Universal Robots PolyScope program: AdientTorsF_Eol20.urp

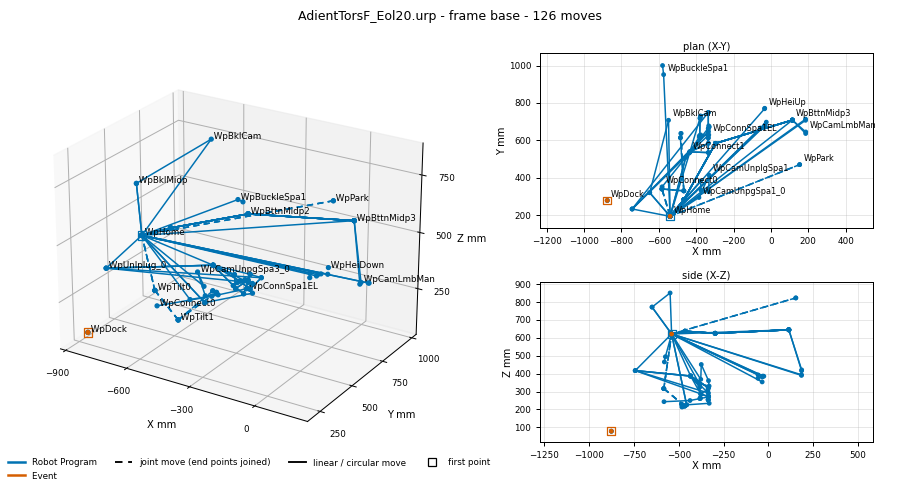
[picture p0: tool path of AdientTorsF_Eol20.urp in frame base, 126 of 179 moves have a stored position in this frame; points joined in program order, loops and branches not executed]
Program AdientTorsF_Eol20 (installation=EOL_20 directory=/programs createdIn=3.5.1 lastSavedIn=5.26.0 robotSerialNumber=20265101888)
Calibrated DH parameters: a=[0.000055, -0.599562, -0.553909, 0.000045, 0.000002, 0]; d=[0.180957, -130.68916, 109.469633, 21.394116, 0.119819, 0.115629]; alpha=[1.570664, -0.000951, 0.006615, 1.571213, -1.569974, 0]; deltaTheta=[0, 0.204436, 5.830565, 0.248193, -0.000001, 0]
InitVariablesNode variables(variable(name=Abort, expression=False), variable(name=AdapterReady, expression=False), variable(name=CMD_Heartbt_i1, expression=0), variable(name=CMD_Program_i1, expression=0), variable(name=CMD_Reserve_i1, expression=0), variable(name=CMD_Timeout_i1, expression=0), variable(name=CamCorrectnOK, expression=0), variable(name=DEBUG, expression=False), variable(name=D_rel, expression=p[0,0,0,0,0,0]), variable(name=EvtBeep, expression=False), variable(name=EvtDock, expression=0), variable(name=Mute, expression=False), variable(name=P_ini, expression=get_actual_tcp_pose()), variable(name=Parking, expression=0), variable(name=ProgExe, expression=0), variable(name=PusherPosFt, expression=0), variable(name=PusherReturn, expression=True), variable(name=STS_Heartbeat, expression=False), variable(name=STS_Progress, expression=0), variable(name=STS_Reservation, expression=0), variable(name=SetCameraProg, expression=0), variable(name=T_KeepReservtn, expression=0), variable(name=Tilt_PV, expression=0))
BeforeStart
  SuppressedNode
    DEBUG := True
  'SW version, to be used to track changes and keep sync of all stations'
  SW_Ver := 1.0
  Folder Scripts [hidden by the author, left out]
  Folder Avoid guidance screen
    Wp := get_actual_tcp_pose()
    MoveJ speed 120 deg/s, acceleration 500 deg/s^2 (useActiveTCP=true optimoveEnabled=false optiMoveSpeed=0.3 optiMoveAcceleration=0.09) feature=Base
      Waypoint Variable (Variable): variable=Wp
  Call GripperOpen
  GoToHome := True
  Script: socket_open("127.0.0.1",30001)
Robot Program (runOnlyOnce=false)
  Folder Execute Program
    Folder Init
      Wait Condition expression=EvtDock≤0
      Folder Verify Adapter ready
        If digital_in[0] or analog_in[3]<(ivGripSensOpen+0.3)
          AdapterReady := False
      Folder Go to home pos automatically
        If GoToHome and  not AdapterReady
          Wait Sleep waitTime=1
          If InRange(P_Flange[0],-1,-0.2) and InRange(P_Flange[1],-0.5,0.5) and InRange(P_Flange[2],0.3,1)
            If AdapterDocked or DEBUG or (analog_in[3]<(ivGripSensOpen+0.3))
              MoveJ speed 120 deg/s, acceleration 500 deg/s^2 (useActiveTCP=false positionType=JointAngles optimoveEnabled=false optiMoveSpeed=0.3 optiMoveAcceleration=0.09) tcp=t0_Flange; feature=Base
                Waypoint WpHome: TCP in base x=-539.74 y=192.879 z=621.496 mm, rx=3.1416 ry=0 rz=0 rad; joints [177.915, -76.399, -107.627, -86.021, 90.391, 88.106] deg
            Else 
              Popup Error (haltProgram=false message=Adapter must be docked inputType=Text)
              Halt
          ElseIf AtParkPos
            MoveJ speed 120 deg/s, acceleration 500 deg/s^2 (useActiveTCP=false positionType=JointAngles optimoveEnabled=false optiMoveSpeed=0.3 optiMoveAcceleration=0.09) tcp=t0_Flange; feature=Base
              Waypoint WpPark: TCP in base x=153.666 y=469.873 z=822.74 mm, rx=-0.0357 ry=3.1413 rz=-0.0002 rad; joints [92.418, -70.926, -90.975, -108.153, 90.407, 181.161] deg
          Else 
            Popup Error (haltProgram=false message=Illegal position. Adjust arm to open space in front of the backrest, or [Move]->[Home] inputType=Text)
            Halt
        GoToHome := False
      If DEBUG
        'Popup window with program selection'
        ProgExe :=  (valueSource=Operator message=Program number? valueType=Integer)
      If ProgExe>0
        Folder Init
          Mute := False
          Wait Condition expression=not GoToHome
          If not In(ProgExe,[11,12,13,14])
            AdapterReady := False
    Folder Programs
      If InRange(ProgExe,1,99)
        Folder Undock
          If In(ProgExe,[11])
            Script: Report(1)
            If not AdapterReady
              Folder AtHome? [hidden by the author, left out]
              If Progress_run() and  not AdapterDocked
                Script: Report(94)
              If Progress_run()
                Folder Undock
                  MoveL speed 1000 mm/s, acceleration 3000 mm/s^2 (useActiveTCP=false optimoveEnabled=false optiMoveSpeed=0.3 optiMoveAcceleration=0.09) tcp=t2_Gripper; feature=Base
                    Call GripperOpenQuick
                    Wp := pose_trans(WpDock, p[0,0.175,-0.1,0,0,0])
                    Waypoint Variable (Variable): motionParameters(blendRadius=0.05); variable=Wp
                    Call GripperOpen
                    Wp := pose_trans(WpDock, p[0,0.075,0.01,0,0,0])
                    Waypoint Variable (Variable): motionParameters(blendRadius=0.01); variable=Wp
                    Wp := pose_trans(WpDock, p[0,0.055,0,0,0,0])
                    Waypoint Variable (Variable): motionParameters(blendRadius=0.01); variable=Wp
                    Waypoint WpDock: TCP in base x=-876.296 y=277.871 z=78.699 mm, rx=1.8725 ry=1.8725 rz=0.5904 rad; joints [172.393, -110.839, -101.123, -92.857, 86.047, -6.096] deg
                    Call GripperClose
                    Wp := pose_trans(WpDock, p[0,0.25,0,0,0,0])
                    Waypoint Variable (Variable): variable=Wp
                  AdapterReady := True
                  Script: Report(50)
            Else 
              Script: Report(50)
        Folder Connect
          If In(ProgExe,[12,13,14])
            Script: Report(1)
            PusherPosDev := 0
            MeasHeight := 0
            If not AdapterReady
              Folder AtHome? [hidden by the author, left out]
              If Progress_run() and  not AdapterDocked
                Script: Report(94)
            If Progress_run()
              Folder Length measure with pusher (mechanical seat)
                If In(ProgExe,[13])
                  Set DigitalOutput pin=Do_PusherReturn; digitalValue=0
                  Set DigitalOutput pin=Do_PusherWork; digitalValue=1
                Else 
                  PusherReturn := True
              Folder Undock
                If not AdapterReady
                  MoveL speed 1000 mm/s, acceleration 3000 mm/s^2 (useActiveTCP=false optimoveEnabled=false optiMoveSpeed=0.3 optiMoveAcceleration=0.09) tcp=t2_Gripper; feature=Base
                    Call GripperOpenQuick
                    Wp := pose_trans(WpDock, p[0,0.175,-0.1,0,0,0])
                    Waypoint Variable (Variable): motionParameters(blendRadius=0.05); variable=Wp
                    Call GripperOpen
                    Wp := pose_trans(WpDock, p[0,0.075,0.01,0,0,0])
                    Waypoint Variable (Variable): motionParameters(blendRadius=0.01); variable=Wp
                    Wp := pose_trans(WpDock, p[0,0.055,0,0,0,0])
                    Waypoint Variable (Variable): motionParameters(blendRadius=0.01); variable=Wp
                    Waypoint WpDock: TCP in base x=-876.296 y=277.871 z=78.699 mm, rx=1.8725 ry=1.8725 rz=0.5904 rad; joints [172.393, -110.839, -101.123, -92.857, 86.047, -6.096] deg
                    Call GripperClose
                    Wp := pose_trans(WpDock, p[0,0.25,0,0,0,0])
                    Waypoint Variable (Variable): variable=Wp
                AdapterReady := False
                Script: Report(2)
              CamCorrection := p[0,0,0,0,0,0]
              SuppressedNode
                Folder Camera
                  MoveL speed 1000 mm/s, acceleration 3000 mm/s^2 (useActiveTCP=false optimoveEnabled=false optiMoveSpeed=0.3 optiMoveAcceleration=0.09) tcp=t0_Flange; feature=Base
                    If In(ProgExe,[12,13])
                      SetCameraProg := 12
                      Waypoint WpCamCon0: motionParameters(blendRadius=0.05); TCP in base x=-326.648 y=291.698 z=338.41 mm, rx=2.1948 ry=2.1949 rz=-0.0575 rad; joints [160.702, -71.24, -141.099, -58.684, 93.132, -18.987] deg
                      Waypoint WpCamConSpa1: TCP in base x=-326.648 y=416.698 z=338.41 mm, rx=2.1948 ry=2.1949 rz=-0.0575 rad; joints [146.583, -82.407, -133.037, -56.241, 92.784, -33.102] deg
                    If In(ProgExe,[14])
                      SetCameraProg := ProgExe
                      Waypoint WpCamCon0: motionParameters(blendRadius=0.05); TCP in base x=-326.648 y=291.698 z=338.41 mm, rx=2.1948 ry=2.1949 rz=-0.0575 rad; joints [160.702, -71.24, -141.099, -58.684, 93.132, -18.987] deg
                      Waypoint WpCamConSpa3: TCP in base x=-370.516 y=382.662 z=354.732 mm, rx=-2.2214 ry=-2.2215 rz=0 rad; joints [153.025, -81.286, -132.366, -56.394, 90.281, -26.621] deg
                  Call CamAcquire
                  CamCorrection := p[CamData[0],CamData[1]*-0.5,CamData[1],0,0,0]
            CamCorrectnOK := ProgExe
            If In(ProgExe,[13])
              Timer (action=Reset) variable=T_Timeout
              Timer (action=Start) variable=T_Timeout
              Wait Condition expression=(PusherPosStable and InRange(PusherPos-ivPusherSeatRef,-15,15)) or T_Timeout>10
              PusherPosDev := PusherPos-ivPusherSeatRef
              If PusherPosStable and InRange(PusherPosDev,-15,15)
                'continue'
              Else 
                CamCorrectnOK := 0
                'CamCorrectionOK is also used as pusher measurement result'
            If Progress_run() and CamCorrectnOK≠ProgExe
              EvtDock := 1
              Wait Condition expression=EvtDock≤0
              Script: Report(91)
            If Progress_run() and ProgExe≟13
              'Wait handle catch done'
              Script: Report(3)
              Timer (action=Reset) variable=T_Timeout
              Timer (action=Start) variable=T_Timeout
              Wait Condition expression=Flags[12] or T_Timeout>10 or DEBUG
              If Flags[12] or DEBUG
                'ok'
              Else 
                Script: Report(98)
            If Progress_run() and  not Di_LiftDown
              EvtDock := 1
              Wait Condition expression=EvtDock≤0
              AdapterReady := False
              Script: Report(92)
            Folder Connect
              If Progress_run()
                Script: Report(4)
                Set NoAction tcp=t2_Gripper
                MoveL speed 1000 mm/s, acceleration 3000 mm/s^2 (useActiveTCP=false optimoveEnabled=false optiMoveSpeed=0.3 optiMoveAcceleration=0.09) tcp=t2_Gripper; feature=Base
                  Waypoint WpConnect0: motionParameters(blendRadius=0.01); TCP in base x=-582.317 y=351.257 z=243.437 mm, rx=-2.2214 ry=-2.2215 rz=0 rad; joints [153.816, -77.664, -139.707, -52.675, 90.266, -25.814] deg; TCP offset x=0 y=-260 z=74 mm, rx=0 ry=0 rz=0 rad
                  Waypoint WpConnect1: TCP in base x=-437.091 y=531.932 z=249.935 mm, rx=3.1416 ry=0 rz=0 rad; joints [167.745, -81.605, -135.899, -52.542, 90.261, 78.118] deg
                  If False
                    Waypoint WpConnSpa1EL: TCP in base x=-332.78 y=629.084 z=270.528 mm, rx=3.1251 ry=-0.0345 rz=0.0169 rad; joints [152.504, -78.36, -135.112, -57.546, 90.839, 64.112] deg
                    Waypoint WpConnSpa1MecTh: TCP in base x=-333.346 y=677.301 z=275.481 mm, rx=3.0512 ry=-0.0001 rz=0 rad; joints [145.822, -81.498, -129.414, -62.023, 94.591, 56.042] deg
                    Waypoint WpConnSpa1Mec: TCP in base x=-335.918 y=624.072 z=312.701 mm, rx=3.0512 ry=-0.0001 rz=0 rad; joints [151.192, -74.921, -130.239, -67.362, 94.873, 61.392] deg
                    Waypoint WpConnSpa3: TCP in base x=-375.972 y=628.734 z=287.575 mm, rx=2.9708 ry=0 rz=0.0001 rad; joints [151.145, -79.992, -126.667, -68.106, 98.894, 61.08] deg
                  If In(ProgExe,[12])
                    Wp := WpConnSpa1EL
                  If In(ProgExe,[13])
                    'adjust angle mechanical'
                    Wp0 := pose_add(WpConnSpa1MecTh,p[0,PusherPosDev/1000,-0.025,0,0,0])
                    Waypoint Variable (Variable): variable=Wp0
                    Force Frame feature=Joint_6_name; selection=[0, 0, 1, 0, 0, 0]; wrench=[0, 0, -30, -0.5, 0, 0]; limitsForce=[0.15, 0.15, 0.1, 0.087266, 1.047198, 1.047198]; limitsMotion=[0.1, 0.1, 0.1, 0.349066, 0.349066, 0.349066]
                      Wait Sleep waitTime=0.5
                    Force Frame feature=Joint_6_name; selection=[0, 0, 1, 0, 0, 0]; wrench=[0, 0, -10, -0.5, 0, 0]; limitsForce=[0.15, 0.15, 0.002, 0.087266, 1.047198, 1.047198]; limitsMotion=[0.1, 0.1, 0.1, 0.349066, 0.349066, 0.349066]
                      Wait Sleep waitTime=0.5
                    Wp := get_actual_tcp_pose()
                    MeasHeight := (Wp[2]-WpConnSpa1MecTh[2])*1000
                    MoveDirectionNode expression=[0.0,1.0,0.2]; feature=Joint_6_name
                      Until DISTANCE (allowActions=false deceleration=3 distanceNodeType=STOP) Distance=0.07; motionParameters(blendRadius=0)
                    Wp := pose_add(WpConnSpa1Mec,p[0,PusherPosDev/1000,0,0,0,0])
                    CorrMechSeat := p[0,0,0,0,0,0]
                    If MeasHeight>0
                      Script: CorrMechSeat[1]=Calibrate(MeasHeight,0,17,0,-7)/1000
                      Script: CorrMechSeat[2]=Calibrate(MeasHeight,0,17,0,26)/1000
                      Script: CorrMechSeat[3]=Calibrate(MeasHeight,0,17,0,-0.129)
                    Else 
                      Script: CorrMechSeat[1]=Calibrate(MeasHeight,-13,0,7,0)/1000
                      Script: CorrMechSeat[2]=Calibrate(MeasHeight,-13,0,-19,0)/1000
                      Script: CorrMechSeat[3]=Calibrate(MeasHeight,-13,0,0.053,0)
                    Wp := pose_add(Wp,CorrMechSeat)
                  If In(ProgExe,[14])
                    Wp := WpConnSpa3
                  Waypoint Variable (Variable): variable=Wp
                Force Frame feature=Joint_6_name; selection=[0, 0, 1, 0, 0, 0]; wrench=[0, 0, -30, 0, 0, 0]; limitsForce=[0.15, 0.15, 0.1, 1.047198, 1.047198, 1.047198]; limitsMotion=[0.1, 0.1, 0.1, 0.349066, 0.349066, 0.349066]
                  Wait Sleep waitTime=1
                Force Frame feature=Joint_6_name; selection=[1, 0, 1, 0, 0, 0]; wrench=[0, 0, -30, 0, 0, 0]; limitsForce=[0.15, 0.15, 0.05, 1.047198, 1.047198, 1.047198]; limitsMotion=[0.1, 0.1, 0.1, 0.349066, 0.349066, 0.349066]
                  Wait Sleep waitTime=0.5
                'position ok, not checked for mechanical seat'
                If InRange(Wp[2]+0.03-P_act[2],-0.015,0.015) or ProgExe≟13
                  'ok'
                Else 
                  EvtDock := 2
                  Wait Condition expression=EvtDock≤0
                  Script: Report(96)
              If Progress_run()
                Force Frame feature=Joint_6_name; selection=[0, 1, 0, 0, 0, 0]; wrench=[0, -60, -10, 0, 0, 0]; limitsForce=[0.15, 0.05, 0.01, 1.047198, 1.047198, 1.047198]; limitsMotion=[0.1, 0.1, 0.1, 0.349066, 0.349066, 0.349066]
                  Wait Sleep waitTime=1
                MoveL speed 1000 mm/s, acceleration 3000 mm/s^2 (useActiveTCP=true optimoveEnabled=false optiMoveSpeed=0.3 optiMoveAcceleration=0.09) feature=Base
                  Wp := pose_trans(P_act, p[0,0.005,0,0,0,0])
                  Waypoint Variable (Variable): variable=Wp
                Call GripperOpen
                Force Frame feature=Joint_6_name; selection=[0, 1, 0, 0, 0, 0]; wrench=[0, -60, -10, 0, 0, 0]; limitsForce=[0.15, 0.1, 0.01, 1.047198, 1.047198, 1.047198]; limitsMotion=[0.1, 0.1, 0.1, 0.349066, 0.349066, 0.349066]
                  Wait Sleep waitTime=1
                  Script: Report(5)
                  MoveL speed 500 mm/s, acceleration 2000 mm/s^2 (useActiveTCP=true optimoveEnabled=false optiMoveSpeed=0.3 optiMoveAcceleration=0.09) feature=Base
                    Wp0 := get_actual_tcp_pose()
                    Wp := pose_trans(Wp0, p[0,0,0,0,0,0.07])
                    Waypoint Variable (Variable): variable=Wp
                    Wp := pose_trans(Wp0, p[0,0,0,0,0,-0.07])
                    Waypoint Variable (Variable): variable=Wp
                    Waypoint Variable (Variable): variable=Wp0
                    Wp := pose_trans(Wp0, p[0,0,0.01,0,0,0])
                    Waypoint Variable (Variable): variable=Wp
                    Waypoint Variable (Variable): variable=Wp0
                MoveL speed 1000 mm/s, acceleration 3000 mm/s^2 (useActiveTCP=true optimoveEnabled=false optiMoveSpeed=0.3 optiMoveAcceleration=0.09) feature=Base
                  Wp0 := get_actual_tcp_pose()
                  Wp := pose_trans(Wp0, p[0,0.015,0,0,0,0])
                  Waypoint Variable (Variable): variable=Wp
                Force Frame feature=Joint_6_name; selection=[0, 1, 0, 0, 0, 0]; wrench=[0, -60, 0, 0, 0, 0]; limitsForce=[0.15, 0.5, 0.15, 1.047198, 1.047198, 1.047198]; limitsMotion=[0.1, 0.1, 0.1, 0.349066, 0.349066, 0.349066]
                  Wait Sleep waitTime=0.5
                Script: Report(6)
                Timer (action=Reset) variable=T_Timeout
                Timer (action=Start) variable=T_Timeout
                Folder Test switch pin, retreat on fail
                  Wait Condition expression=Flags[0] or T_Timeout>10 or DEBUG
                  If not Flags[0] and  not DEBUG
                    EvtDock := 2
                    Wait Condition expression=EvtDock≤0
                    Script: Report(95)
            If Progress_run()
              MoveL speed 1000 mm/s, acceleration 3000 mm/s^2 (useActiveTCP=false optimoveEnabled=false optiMoveSpeed=0.3 optiMoveAcceleration=0.09) tcp=t0_Flange; feature=Base
                Set NoAction tcp=t0_Flange
                P_act := get_actual_tcp_pose()
                Wp := pose_trans(P_act, p[0,0.1,0,0,0,0])
                Waypoint Variable (Variable): motionParameters(blendRadius=0.05); variable=Wp
                Wp := pose_trans(Wp, p[-0.15,0.1,-0.2,0,0.5,0])
                Waypoint Variable (Variable): motionParameters(blendRadius=0.05); variable=Wp
                Waypoint WpHome: TCP in base x=-539.74 y=192.879 z=621.496 mm, rx=3.1416 ry=0 rz=0 rad; joints [177.915, -76.399, -107.627, -86.021, 90.391, 88.106] deg
              Script: Report(50)
        Folder Buckle
          If In(ProgExe,[15,16])
            Script: Report(1)
            Folder AtHome? [hidden by the author, left out]
            If Progress_run() and  not Di_SBR_X_Wp
              Script: Report(92)
            If Progress_run()
              Call GripperCloseQuick
              Folder Camera
                SetCameraProg := ProgExe
                MoveL speed 1000 mm/s, acceleration 3000 mm/s^2 (useActiveTCP=false optimoveEnabled=false optiMoveSpeed=0.3 optiMoveAcceleration=0.09) tcp=t0_Flange; feature=Base
                  Waypoint WpBklCam: TCP in base x=-548.167 y=707.316 z=850.607 mm, rx=-1.8029 ry=-0.697 rz=1.8635 rad; joints [133.218, -113.859, -67.455, 3.142, 139.231, 51.988] deg
                Call GripperClose
                Call CamAcquire
                Call CamCalculateCorectnPlane
                If CamCorrectnOK≟ProgExe and InRange(CamCorrection[1],-0.05,0.05) and InRange(CamCorrection[2],-0.03,0.03)
                  'empty'
                Else 
                  CamCorrectnOK := 0
                  MoveL speed 1000 mm/s, acceleration 3000 mm/s^2 (useActiveTCP=false optimoveEnabled=false optiMoveSpeed=0.3 optiMoveAcceleration=0.09) tcp=t0_Flange; feature=Base
                    Waypoint WpBklMidp: motionParameters(blendRadius=0.05); TCP in base x=-648.886 y=319.496 z=771.546 mm, rx=3.1416 ry=0 rz=0 rad; joints [167.64, -91.713, -78.917, -99.416, 90.395, 77.75] deg
                    Waypoint WpHome: TCP in base x=-539.74 y=192.879 z=621.496 mm, rx=3.1416 ry=0 rz=0 rad; joints [177.915, -76.399, -107.627, -86.021, 90.391, 88.106] deg
                  Script: Report(91)
              If CamCorrectnOK≟ProgExe
                Folder Insert
                  MoveL speed 1000 mm/s, acceleration 3000 mm/s^2 (useActiveTCP=false optimoveEnabled=false optiMoveSpeed=0.3 optiMoveAcceleration=0.09) tcp=t3_Blade; feature=Base
                    If False
                      'must be set with blade ca one half into buckle slot'
                      Waypoint WpBuckleSpa1: TCP in base x=-574.481 y=951.559 z=494.56 mm, rx=-2.7053 ry=0 rz=0 rad; joints [140.754, -127.124, -55.008, -71.575, 71.185, 48.273] deg; TCP offset x=134 y=-56 z=118 mm, rx=0 ry=0 rz=0 rad
                      Waypoint WpBuckleSpa3: TCP in base x=-580.216 y=1000.227 z=465.338 mm, rx=-2.606 ry=0.0419 rz=-0.222 rad; joints [140.4, -134.437, -48.452, -74.762, 61.024, 49.269] deg
                    If ProgExe≟15
                      Wp := WpBuckleSpa1
                    If ProgExe≟16
                      Wp := WpBuckleSpa3
                    Wp0 := pose_trans(Wp,p[0,0,-0.02,0,0,0])
                    Wp0 := pose_add(Wp0,Base_w_correctn)
                    Waypoint Variable (Variable): variable=Wp0
                  Script: Report(5)
                  Timer (action=Reset) variable=T_Timeout
                  Timer (action=Start) variable=T_Timeout
                  Wait Condition expression=Flags[8] or Abort or DEBUG  or T_Timeout>25
                  If Flags[8] or DEBUG
                    Script: Report(6)
                    Set NoAction tcp=t3_Blade
                    Force Frame feature=Joint_6_name; selection=[0, 0, 1, 0, 0, 0]; wrench=[0, 0, 15, 0, 0, 0]; limitsForce=[0.15, 0.15, 0.15, 1.047198, 1.047198, 1.047198]; limitsMotion=[0.1, 0.1, 0.1, 0.349066, 0.349066, 0.349066]
                      Wait Sleep waitTime=1
                    If not Flags[9] and  not Abort
                      MoveL speed 50 mm/s, acceleration 500 mm/s^2 (useActiveTCP=false optimoveEnabled=false optiMoveSpeed=0.3 optiMoveAcceleration=0.09) tcp=t3_Blade; feature=Base
                        Waypoint Variable (Variable): variable=Wp
                      Force Frame feature=Joint_6_name; selection=[1, 1, 1, 0, 0, 0]; wrench=[0, 0, 50, 0, 0, 0]; limitsForce=[0.15, 0.15, 0.25, 1.047198, 1.047198, 1.047198]; limitsMotion=[0.1, 0.1, 0.1, 0.349066, 0.349066, 0.349066]
                        Wait Sleep waitTime=1.5
                    If not Flags[9] and  not Abort
                      MoveL speed 50 mm/s, acceleration 500 mm/s^2 (useActiveTCP=false optimoveEnabled=false optiMoveSpeed=0.3 optiMoveAcceleration=0.09) tcp=t3_Blade; feature=Base
                        Waypoint Variable (Variable): variable=Wp
                      Force Frame feature=Joint_6_name; selection=[1, 1, 1, 0, 0, 0]; wrench=[0, 0, 50, 0, 0, 0]; limitsForce=[0.15, 0.15, 0.25, 1.047198, 1.047198, 1.047198]; limitsMotion=[0.1, 0.1, 0.1, 0.349066, 0.349066, 0.349066]
                        Wait Sleep waitTime=1.5
                    If not Flags[9] and  not Abort
                      MoveL speed 50 mm/s, acceleration 500 mm/s^2 (useActiveTCP=false optimoveEnabled=false optiMoveSpeed=0.3 optiMoveAcceleration=0.09) tcp=t3_Blade; feature=Base
                        Waypoint Variable (Variable): variable=Wp
                      Force Frame feature=Joint_6_name; selection=[1, 1, 1, 0, 0, 0]; wrench=[0, 0, 50, 0, 0, 0]; limitsForce=[0.15, 0.15, 0.25, 1.047198, 1.047198, 1.047198]; limitsMotion=[0.1, 0.1, 0.1, 0.349066, 0.349066, 0.349066]
                        Wait Sleep waitTime=1.5
                  MoveL speed 1000 mm/s, acceleration 3000 mm/s^2 (useActiveTCP=false optimoveEnabled=false optiMoveSpeed=0.3 optiMoveAcceleration=0.09) tcp=t3_Blade; feature=Base
                    Waypoint Variable (Variable): variable=Wp
                    MoveDirectionNode (selectedDirection=ZMinus) feature=Joint_6_name
                      Until DISTANCE (allowActions=false deceleration=3 distanceNodeType=STOP) Distance=0.02; motionParameters(blendRadius=0)
                  MoveL speed 1000 mm/s, acceleration 3000 mm/s^2 (useActiveTCP=false optimoveEnabled=false optiMoveSpeed=0.3 optiMoveAcceleration=0.09) tcp=t0_Flange; feature=Base
                    Waypoint WpBklMidp: motionParameters(blendRadius=0.05); TCP in base x=-648.886 y=319.496 z=771.546 mm, rx=3.1416 ry=0 rz=0 rad; joints [167.64, -91.713, -78.917, -99.416, 90.395, 77.75] deg
                    Waypoint WpHome: TCP in base x=-539.74 y=192.879 z=621.496 mm, rx=3.1416 ry=0 rz=0 rad; joints [177.915, -76.399, -107.627, -86.021, 90.391, 88.106] deg
                  If Progress_check()≥6
                    Script: Report(50)
                  Else 
                    Script: Report(95)
        Folder Disconnect
          If In(ProgExe,[21,22,23])
            Script: Report(1)
            Folder AtHome? [hidden by the author, left out]
            If Progress_run()
              If In(ProgExe,[21])
                SetCameraProg := ProgExe
                MoveL speed 1000 mm/s, acceleration 3000 mm/s^2 (useActiveTCP=false optimoveEnabled=false optiMoveSpeed=0.3 optiMoveAcceleration=0.09) tcp=t0_Flange; feature=Base
                  Waypoint WpCamUnpgSpa1_0: motionParameters(blendRadius=0.05); TCP in base x=-385.489 y=293.712 z=344.085 mm, rx=2.1641 ry=2.1642 rz=-0.1205 rad; joints [162.074, -77.174, -136.372, -58.433, 96.359, -17.691] deg
                  Waypoint WpCamUnplgSpa1: TCP in base x=-330.386 y=412.98 z=330.769 mm, rx=2.1642 ry=2.1642 rz=-0.1205 rad; joints [146.528, -83.262, -132.856, -57.421, 95.6, -33.289] deg
              If In(ProgExe,[22])
                SetCameraProg := ProgExe
                MoveL speed 1000 mm/s, acceleration 3000 mm/s^2 (useActiveTCP=false optimoveEnabled=false optiMoveSpeed=0.3 optiMoveAcceleration=0.09) tcp=t0_Flange; feature=Base
                  Waypoint WpCamUnplgSpa1M: TCP in base x=-333.812 y=324.612 z=360.892 mm, rx=2.1642 ry=2.1642 rz=-0.1205 rad; joints [156.073, -73.679, -136.623, -62.306, 96.141, -23.739] deg
              If In(ProgExe,[23])
                SetCameraProg := ProgExe
                MoveL speed 1000 mm/s, acceleration 3000 mm/s^2 (useActiveTCP=false optimoveEnabled=false optiMoveSpeed=0.3 optiMoveAcceleration=0.09) tcp=t0_Flange; feature=Base
                  Waypoint WpCamUnpgSpa3_0: motionParameters(blendRadius=0.05); TCP in base x=-374.135 y=332.475 z=451.177 mm, rx=2.1642 ry=2.1642 rz=-0.1205 rad; joints [157.169, -73.07, -127.046, -72.385, 96.229, -22.692] deg
                  Waypoint WpCamUnpgSpa3: TCP in base x=-376.961 y=382.567 z=368.205 mm, rx=2.1236 ry=2.1236 rz=-0.1987 rad; joints [151.263, -82.063, -129.1, -64.018, 99.681, -28.849] deg
              Call CamAcquire
              Call CamCalculateCorectnPlane
            If Progress_run() and CamCorrectnOK≠ProgExe
              MoveL speed 1000 mm/s, acceleration 3000 mm/s^2 (useActiveTCP=false optimoveEnabled=false optiMoveSpeed=0.3 optiMoveAcceleration=0.09) tcp=t0_Flange; feature=Base
                Waypoint WpHome: TCP in base x=-539.74 y=192.879 z=621.496 mm, rx=3.1416 ry=0 rz=0 rad; joints [177.915, -76.399, -107.627, -86.021, 90.391, 88.106] deg
              Script: Report(91)
            If Progress_run()
              Call GripperOpenQuick
              Folder Disconnect
                If In(ProgExe,[21])
                  MoveL speed 1000 mm/s, acceleration 3000 mm/s^2 (useActiveTCP=false optimoveEnabled=false optiMoveSpeed=0.3 optiMoveAcceleration=0.09) tcp=t2_Gripper; feature=Base_w_correctn
                    Waypoint WpUnlplug_0: motionParameters(blendRadius=0.05); TCP in base x=-742.864 y=232.307 z=416.977 mm, rx=2.2214 ry=2.2214 rz=0 rad; joints [173.149, -74.838, -122.091, -73.118, 90.357, -6.582] deg; TCP offset x=0 y=-260 z=74 mm, rx=0 ry=0 rz=0 rad
                    Call GripperOpen
                    Waypoint WpUnplug_1: motionParameters(blendRadius=0.05); TCP in base x=-433.594 y=537.985 z=386.664 mm, rx=3.1416 ry=0 rz=0 rad; joints [166.968, -73.547, -126.184, -70.315, 90.348, 77.251] deg
                    Waypoint WpUnplug1_15: motionParameters(blendRadius=0.05); TCP in base x=-335.185 y=584.129 z=321.99 mm, rx=2.6768 ry=0 rz=0 rad; joints [145.854, -75.949, -117.78, -91.984, 112.189, 52.946] deg
                    Waypoint WpUnplug1_2: motionParameters(blendRadius=0.05); TCP in base x=-335.446 y=662.579 z=254.257 mm, rx=2.6768 ry=0 rz=0 rad; joints [139.434, -84.88, -117.162, -86.002, 110.307, 46.418] deg
                    Waypoint WpUnplug1_3: TCP in base x=-335.273 y=749.502 z=272.417 mm, rx=3.0593 ry=-0.0005 rz=0.0001 rad; joints [140.09, -87.914, -124.299, -60.846, 93.913, 50.349] deg
                If In(ProgExe,[22])
                  MoveL speed 1000 mm/s, acceleration 3000 mm/s^2 (useActiveTCP=false optimoveEnabled=false optiMoveSpeed=0.3 optiMoveAcceleration=0.09) tcp=t2_Gripper; feature=Base_w_correctn
                    Waypoint WpUnlplug_0: motionParameters(blendRadius=0.05); TCP in base x=-742.864 y=232.307 z=416.977 mm, rx=2.2214 ry=2.2214 rz=0 rad; joints [173.149, -74.838, -122.091, -73.118, 90.357, -6.582] deg
                    Call GripperOpen
                    Waypoint WpUnplug_1: motionParameters(blendRadius=0.05); TCP in base x=-433.594 y=537.985 z=386.664 mm, rx=3.1416 ry=0 rz=0 rad; joints [166.968, -73.547, -126.184, -70.315, 90.348, 77.251] deg
                    Waypoint WpUnplug_1_1M: motionParameters(blendRadius=0.05); TCP in base x=-335.185 y=534.129 z=321.99 mm, rx=2.6768 ry=0 rz=0 rad; joints [150.71, -71.65, -121.165, -90.956, 113.427, 58.032] deg; TCP offset x=0 y=-260 z=74 mm, rx=0 ry=0 rz=0 rad
                    Waypoint WpUnplug1_2M: motionParameters(blendRadius=0.05); TCP in base x=-335.446 y=612.579 z=254.257 mm, rx=2.6768 ry=0 rz=0 rad; joints [143.376, -80.619, -121.11, -84.903, 111.483, 50.441] deg; TCP offset x=0 y=-260 z=74 mm, rx=0 ry=0 rz=0 rad
                    Waypoint WpUnplg1_3M: TCP in base x=-335.273 y=646.793 z=292.13 mm, rx=2.9682 ry=-0.0005 rz=0.0001 rad; joints [147.069, -78.306, -127.241, -69.901, 98.673, 56.974] deg; TCP offset x=0 y=-260 z=74 mm, rx=0 ry=0 rz=0 rad
                    SuppressedNode
                      Waypoint Waypoint_1: TCP in base x=-335.273 y=649.502 z=297.176 mm, rx=3.0593 ry=-0.0005 rz=0.0001 rad; joints [148.743, -77.933, -130.038, -64.507, 94.352, 58.989] deg
                If In(ProgExe,[23])
                  MoveL speed 1000 mm/s, acceleration 3000 mm/s^2 (useActiveTCP=false optimoveEnabled=false optiMoveSpeed=0.3 optiMoveAcceleration=0.09) tcp=t2_Gripper; feature=Base_w_correctn
                    Waypoint WpUnlplug_0: motionParameters(blendRadius=0.05); TCP in base x=-742.864 y=232.307 z=416.977 mm, rx=2.2214 ry=2.2214 rz=0 rad; joints [173.149, -74.838, -122.091, -73.118, 90.357, -6.582] deg
                    Call GripperOpen
                    Waypoint WpUnplug_1: motionParameters(blendRadius=0.05); TCP in base x=-433.594 y=537.985 z=386.664 mm, rx=3.1416 ry=0 rz=0 rad; joints [166.968, -73.547, -126.184, -70.315, 90.348, 77.251] deg
                    Waypoint WpUnplg3_2: motionParameters(blendRadius=0.05); TCP in base x=-382.207 y=617.524 z=326.263 mm, rx=2.948 ry=0 rz=0 rad; joints [152.036, -77.933, -123.356, -73.967, 100.146, 61.843] deg
                    Waypoint WpUnplg3_3: motionParameters(blendRadius=0.014); TCP in base x=-381.485 y=624.575 z=260.915 mm, rx=2.948 ry=0 rz=0 rad; joints [151.318, -81.621, -127.658, -66.093, 100.047, 61.163] deg
                    Waypoint WpUnplg3_4: motionParameters(blendRadius=0.023); TCP in base x=-379.373 y=718.034 z=263.548 mm, rx=2.948 ry=0 rz=0 rad; joints [143.235, -88.587, -120.8, -67.307, 99.196, 53.013] deg
                    Waypoint WpUnplg3_5: TCP in base x=-376.755 y=729.692 z=285.292 mm, rx=2.948 ry=0 rz=0 rad; joints [142.211, -88.242, -118.628, -69.985, 99.086, 51.969] deg
                Script: Report(20)
                Wait Condition expression=Flags[7] or DEBUG
              EvtDock := 2
              Wait Condition expression=EvtDock≤0
              If EvtDock<0
                If In(ProgExe,[21])
                  MoveL speed 1000 mm/s, acceleration 3000 mm/s^2 (useActiveTCP=false optimoveEnabled=false optiMoveSpeed=0.3 optiMoveAcceleration=0.09) tcp=t2_Gripper; feature=Base_w_correctn
                    Waypoint WpUnplug1_3: TCP in base x=-335.273 y=749.502 z=272.417 mm, rx=3.0593 ry=-0.0005 rz=0.0001 rad; joints [140.09, -87.914, -124.299, -60.846, 93.913, 50.349] deg
                    Waypoint WpUnplug1_2: TCP in base x=-335.446 y=662.579 z=254.257 mm, rx=2.6768 ry=0 rz=0 rad; joints [139.434, -84.88, -117.162, -86.002, 110.307, 46.418] deg
                    Waypoint WpUnplug1_15: TCP in base x=-335.185 y=584.129 z=321.99 mm, rx=2.6768 ry=0 rz=0 rad; joints [145.854, -75.949, -117.78, -91.984, 112.189, 52.946] deg
                    Waypoint WpUnplug_1: TCP in base x=-433.594 y=537.985 z=386.664 mm, rx=3.1416 ry=0 rz=0 rad; joints [166.968, -73.547, -126.184, -70.315, 90.348, 77.251] deg
                    SuppressedNode
                      Waypoint WpUnlplug_0: motionParameters(blendRadius=0.05); TCP in base x=-742.864 y=232.307 z=416.977 mm, rx=2.2214 ry=2.2214 rz=0 rad; joints [173.149, -74.838, -122.091, -73.118, 90.357, -6.582] deg
                If In(ProgExe,[22])
                  MoveL speed 1000 mm/s, acceleration 3000 mm/s^2 (useActiveTCP=false optimoveEnabled=false optiMoveSpeed=0.3 optiMoveAcceleration=0.09) tcp=t2_Gripper; feature=Base_w_correctn
                    Waypoint WpUnplg1_3M: TCP in base x=-335.273 y=646.793 z=292.13 mm, rx=2.9682 ry=-0.0005 rz=0.0001 rad; joints [147.069, -78.306, -127.241, -69.901, 98.673, 56.974] deg
                    Waypoint WpUnplug1_2M: TCP in base x=-335.446 y=612.579 z=254.257 mm, rx=2.6768 ry=0 rz=0 rad; joints [143.376, -80.619, -121.11, -84.903, 111.483, 50.441] deg; TCP offset x=0 y=-260 z=74 mm, rx=0 ry=0 rz=0 rad
                    Waypoint WpUnplug_1_1M: TCP in base x=-335.185 y=534.129 z=321.99 mm, rx=2.6768 ry=0 rz=0 rad; joints [150.71, -71.65, -121.165, -90.956, 113.427, 58.032] deg; TCP offset x=0 y=-260 z=74 mm, rx=0 ry=0 rz=0 rad
                    Waypoint WpUnplug_1: TCP in base x=-433.594 y=537.985 z=386.664 mm, rx=3.1416 ry=0 rz=0 rad; joints [166.968, -73.547, -126.184, -70.315, 90.348, 77.251] deg; TCP offset x=0 y=-260 z=74 mm, rx=0 ry=0 rz=0 rad
                    SuppressedNode
                      Waypoint WpUnlplug_0: motionParameters(blendRadius=0.05); TCP in base x=-742.864 y=232.307 z=416.977 mm, rx=2.2214 ry=2.2214 rz=0 rad; joints [173.149, -74.838, -122.091, -73.118, 90.357, -6.582] deg
                If In(ProgExe,[23])
                  MoveL speed 1000 mm/s, acceleration 3000 mm/s^2 (useActiveTCP=false optimoveEnabled=false optiMoveSpeed=0.3 optiMoveAcceleration=0.09) tcp=t2_Gripper; feature=Base_w_correctn
                    Waypoint WpUnplg3_5: TCP in base x=-376.755 y=729.692 z=285.292 mm, rx=2.948 ry=0 rz=0 rad; joints [142.211, -88.242, -118.628, -69.985, 99.086, 51.969] deg
                    Waypoint WpUnplg3_4: TCP in base x=-379.373 y=718.034 z=263.548 mm, rx=2.948 ry=0 rz=0 rad; joints [143.235, -88.587, -120.8, -67.307, 99.196, 53.013] deg
                    Waypoint WpUnplg3_3: TCP in base x=-381.485 y=624.575 z=260.915 mm, rx=2.948 ry=0 rz=0 rad; joints [151.318, -81.621, -127.658, -66.093, 100.047, 61.163] deg
                    Waypoint WpUnplg3_2: motionParameters(blendRadius=0.05); TCP in base x=-382.207 y=617.524 z=326.263 mm, rx=2.948 ry=0 rz=0 rad; joints [152.036, -77.933, -123.356, -73.967, 100.146, 61.843] deg
                    Waypoint WpUnplug_1: motionParameters(blendRadius=0.05); TCP in base x=-433.594 y=537.985 z=386.664 mm, rx=3.1416 ry=0 rz=0 rad; joints [166.968, -73.547, -126.184, -70.315, 90.348, 77.251] deg
                    SuppressedNode
                      Waypoint WpUnlplug_0: motionParameters(blendRadius=0.05); TCP in base x=-742.864 y=232.307 z=416.977 mm, rx=2.2214 ry=2.2214 rz=0 rad; joints [173.149, -74.838, -122.091, -73.118, 90.357, -6.582] deg
                MoveL speed 1000 mm/s, acceleration 3000 mm/s^2 (useActiveTCP=false optimoveEnabled=false optiMoveSpeed=0.3 optiMoveAcceleration=0.09) tcp=t0_Flange; feature=Base
                  Waypoint WpHome: TCP in base x=-539.74 y=192.879 z=621.496 mm, rx=3.1416 ry=0 rz=0 rad; joints [177.915, -76.399, -107.627, -86.021, 90.391, 88.106] deg
                Script: Report(97)
            If Progress_run()
              Script: Report(50)
        Folder Buttons
          If In(ProgExe,[31,32,34])
            Script: Report(1)
            Folder AtHome? [hidden by the author, left out]
            Folder Camera
              If Progress_run()
                If In(ProgExe,[31,32])
                  SetCameraProg := 32
                  MeasHeight := 0
                If In(ProgExe,[34])
                  SetCameraProg := 34
                MoveL speed 1000 mm/s, acceleration 3000 mm/s^2 (useActiveTCP=false optimoveEnabled=false optiMoveSpeed=0.3 optiMoveAcceleration=0.09) tcp=t0_Flange; feature=Base
                  Waypoint WpBttnMidp1: motionParameters(blendRadius=0.1); TCP in base x=-465.361 y=283.426 z=636.73 mm, rx=-2.2214 ry=2.2214 rz=0 rad; joints [167.185, -73.405, -108.257, -88.385, 90.398, 167.36] deg
                  Waypoint WpBttnMidp2: motionParameters(blendRadius=0.1); TCP in base x=-296.641 y=583.561 z=625.265 mm, rx=-1.2596 ry=2.878 rz=0 rad; joints [132.275, -84.542, -100.549, -84.955, 90.381, 175.201] deg
                  Waypoint WpBttnMidp3: motionParameters(blendRadius=0.1); TCP in base x=114.747 y=708.142 z=644.758 mm, rx=0 ry=3.1416 rz=0 rad; joints [94.755, -90.505, -92.903, -86.639, 90.379, 184.947] deg; TCP offset x=0 y=0 z=0 mm, rx=0 ry=0 rz=0 rad
                  If In(ProgExe,[34])
                    If False
                      Waypoint WpCamLmbMan: TCP in base x=186.376 y=644.645 z=421 mm, rx=0.3238 ry=3.0539 rz=-0.0115 rad; joints [89.517, -91.508, -115.089, -64.291, 86.326, 191.973] deg; TCP offset x=0 y=0 z=0 mm, rx=0 ry=0 rz=0 rad
                    Wp := pose_add(WpCamLmbMan,p[0,0,MeasHeight/1000,0,0,0])
                    Waypoint Variable (Variable): variable=Wp
                  Else 
                    Waypoint WpCamLmbEL: TCP in base x=185.817 y=636.329 z=416.403 mm, rx=0.3238 ry=3.0539 rz=-0.0115 rad; joints [89.561, -90.94, -116.187, -63.764, 86.325, 192.02] deg
                Call CamAcquire
                Script: CamData[1]=CamData[1]-MeasHeight/1000
                Call CamCalculateCorectnPlane
            If Progress_run() and CamCorrectnOK≠ProgExe
              MoveL speed 1000 mm/s, acceleration 3000 mm/s^2 (useActiveTCP=false optimoveEnabled=false optiMoveSpeed=0.3 optiMoveAcceleration=0.09) tcp=t0_Flange; feature=Base
                Waypoint WpBttnMidp3: motionParameters(blendRadius=0.1); TCP in base x=114.747 y=708.142 z=644.758 mm, rx=0 ry=3.1416 rz=0 rad; joints [94.755, -90.505, -92.903, -86.639, 90.379, 184.947] deg; TCP offset x=0 y=0 z=0 mm, rx=0 ry=0 rz=0 rad
                Waypoint WpBttnMidp2: motionParameters(blendRadius=0.1); TCP in base x=-296.641 y=583.561 z=625.265 mm, rx=-1.2596 ry=2.878 rz=0 rad; joints [132.275, -84.542, -100.549, -84.955, 90.381, 175.201] deg
                Waypoint WpBttnMidp1: motionParameters(blendRadius=0.1); TCP in base x=-465.361 y=283.426 z=636.73 mm, rx=-2.2214 ry=2.2214 rz=0 rad; joints [167.185, -73.405, -108.257, -88.385, 90.398, 167.36] deg
                Waypoint WpHome: TCP in base x=-539.74 y=192.879 z=621.496 mm, rx=3.1416 ry=0 rz=0 rad; joints [177.915, -76.399, -107.627, -86.021, 90.391, 88.106] deg
              Script: Report(91)
            Folder Lumbar
              If Progress_run()
                If In(ProgExe,[31,32])
                  Timer (action=Reset) variable=T_Timeout
                  Timer (action=Start) variable=T_Timeout
                  Script: Report(12)
                  Wait Condition expression=Flags[2] or T_Timeout>60 or DEBUG or Abort
                  If Flags[2] or DEBUG
                    MoveL speed 1000 mm/s, acceleration 3000 mm/s^2 (useActiveTCP=false optimoveEnabled=false optiMoveSpeed=0.3 optiMoveAcceleration=0.09) tcp=t4_Finger; feature=Base
                      Folder Press FW
                        If False
                          Waypoint WpLmbFwEL: TCP in base x=-33.633 y=677.236 z=382.161 mm, rx=0.3312 ry=3.1241 rz=0 rad; joints [93.201, -94.299, -108.853, -66.894, 90.316, 195.61] deg; TCP offset x=159 y=-58 z=70 mm, rx=0 ry=0 rz=0 rad
                        Wp := pose_trans(WpLmbFwEL, CamCorrection)
                        Waypoint Variable (Variable): variable=Wp
                        Force Frame feature=Joint_6_name; selection=[1, 0, 0, 0, 0, 0]; wrench=[20, 10, -20, 0, 0, 0]; limitsForce=[0.05, 0.01, 0.05, 1.047198, 1.047198, 1.047198]; limitsMotion=[0.1, 0.1, 0.1, 0.349066, 0.349066, 0.349066]
                          Wait Sleep waitTime=0.7
                        ButtonPos := get_actual_tcp_pose()
                        Waypoint Variable (Variable): variable=Wp
                    Script: Report(3)
                  Else 
                    MoveL speed 1000 mm/s, acceleration 3000 mm/s^2 (useActiveTCP=false optimoveEnabled=false optiMoveSpeed=0.3 optiMoveAcceleration=0.09) tcp=t0_Flange; feature=Base
                      Waypoint WpBttnMidp3: motionParameters(blendRadius=0.1); TCP in base x=114.747 y=708.142 z=644.758 mm, rx=0 ry=3.1416 rz=0 rad; joints [94.755, -90.505, -92.903, -86.639, 90.379, 184.947] deg; TCP offset x=0 y=0 z=0 mm, rx=0 ry=0 rz=0 rad
                      Waypoint WpBttnMidp2: motionParameters(blendRadius=0.1); TCP in base x=-296.641 y=583.561 z=625.265 mm, rx=-1.2596 ry=2.878 rz=0 rad; joints [132.275, -84.542, -100.549, -84.955, 90.381, 175.201] deg
                      Waypoint WpBttnMidp1: motionParameters(blendRadius=0.1); TCP in base x=-465.361 y=283.426 z=636.73 mm, rx=-2.2214 ry=2.2214 rz=0 rad; joints [167.185, -73.405, -108.257, -88.385, 90.398, 167.36] deg
                      Waypoint WpHome: TCP in base x=-539.74 y=192.879 z=621.496 mm, rx=3.1416 ry=0 rz=0 rad; joints [177.915, -76.399, -107.627, -86.021, 90.391, 88.106] deg
                    Script: Report(95)
            Folder Multiring
              If Progress_run()
                If In(ProgExe,[32])
                  Timer (action=Reset) variable=T_Timeout
                  Timer (action=Start) variable=T_Timeout
                  Script: Report(11)
                  Wait Condition expression=Flags[1] or T_Timeout>60 or DEBUG or Abort
                  If Flags[1] or DEBUG
                    MoveL speed 1000 mm/s, acceleration 3000 mm/s^2 (useActiveTCP=false optimoveEnabled=false optiMoveSpeed=0.3 optiMoveAcceleration=0.09) tcp=t4_Finger; feature=Base
                      If False
                        Waypoint WpMultiringHi: TCP in base x=-56.848 y=665.442 z=392.873 mm, rx=0.3312 ry=3.1241 rz=0 rad; joints [95.214, -92.416, -109.702, -67.928, 90.322, 197.618] deg; TCP offset x=159 y=-58 z=70 mm, rx=0 ry=0 rz=0 rad
                        Waypoint WpMutiringLo: TCP in base x=-57.199 y=664.623 z=373.904 mm, rx=-0.3307 ry=-3.1199 rz=0.0014 rad; joints [95.181, -93.124, -111.101, -65.823, 90.559, 197.596] deg
                      Folder Press up
                        Wp0 := pose_add(WpMutiringLo,Base_w_correctn)
                        Wp0 := pose_trans(Wp0, p[-0.02,0,0,0,0,0])
                        Wp := Wp0
                        Script: Wp[0]=ButtonPos[0]-0.01
                        Waypoint Variable (Variable): variable=Wp0
                        Waypoint Variable (Variable): variable=Wp
                        Set NoAction tcp=t4_Finger
                        Force Frame feature=Joint_6_name; selection=[0, 1, 1, 0, 0, 0]; wrench=[10, 20, -20, 0, 0, 0]; limitsForce=[0.01, 0.01, 0.025, 1.047198, 1.047198, 1.047198]; limitsMotion=[0.1, 0.1, 0.1, 0.349066, 0.349066, 0.349066]
                          Wait Sleep waitTime=1
                        Waypoint Variable (Variable): variable=Wp0
                      Folder Press down
                        Wp0 := pose_add(WpMultiringHi,Base_w_correctn)
                        Wp0 := pose_trans(Wp0, p[-0.02,0,0,0,0,0])
                        Wp := Wp0
                        Script: Wp[0]=ButtonPos[0]
                        Script: Wp[0]=ButtonPos[0]-0.01
                        Waypoint Variable (Variable): variable=Wp0
                        Waypoint Variable (Variable): variable=Wp
                        Set NoAction tcp=t4_Finger
                        Force Frame feature=Joint_6_name; selection=[0, 1, 1, 0, 0, 0]; wrench=[10, 20, 20, 0, 0, 0]; limitsForce=[0.01, 0.01, 0.05, 1.047198, 1.047198, 1.047198]; limitsMotion=[0.1, 0.1, 0.1, 0.349066, 0.349066, 0.349066]
                          Wait Sleep waitTime=1
                        Waypoint Variable (Variable): variable=Wp0
                    Script: Report(2)
                  Else 
                    MoveL speed 1000 mm/s, acceleration 3000 mm/s^2 (useActiveTCP=false optimoveEnabled=false optiMoveSpeed=0.3 optiMoveAcceleration=0.09) tcp=t0_Flange; feature=Base
                      Waypoint WpBttnMidp3: motionParameters(blendRadius=0.1); TCP in base x=114.747 y=708.142 z=644.758 mm, rx=0 ry=3.1416 rz=0 rad; joints [94.755, -90.505, -92.903, -86.639, 90.379, 184.947] deg; TCP offset x=0 y=0 z=0 mm, rx=0 ry=0 rz=0 rad
                      Waypoint WpBttnMidp2: motionParameters(blendRadius=0.1); TCP in base x=-296.641 y=583.561 z=625.265 mm, rx=-1.2596 ry=2.878 rz=0 rad; joints [132.275, -84.542, -100.549, -84.955, 90.381, 175.201] deg
                      Waypoint WpBttnMidp1: motionParameters(blendRadius=0.1); TCP in base x=-465.361 y=283.426 z=636.73 mm, rx=-2.2214 ry=2.2214 rz=0 rad; joints [167.185, -73.405, -108.257, -88.385, 90.398, 167.36] deg
                      Waypoint WpHome: TCP in base x=-539.74 y=192.879 z=621.496 mm, rx=3.1416 ry=0 rz=0 rad; joints [177.915, -76.399, -107.627, -86.021, 90.391, 88.106] deg
                    Script: Report(95)
            Folder 2W LMB FW
              If Progress_run()
                If In(ProgExe,[34])
                  SetCameraProg := 35
                  Timer (action=Reset) variable=T_Timeout
                  Timer (action=Start) variable=T_Timeout
                  Script: Report(13)
                  Wait Condition expression=Flags[3] or T_Timeout>60 or DEBUG or Abort
                  If Flags[3] or DEBUG
                    MoveL speed 1000 mm/s, acceleration 3000 mm/s^2 (useActiveTCP=false optimoveEnabled=false optiMoveSpeed=0.3 optiMoveAcceleration=0.09) tcp=t4_Finger; feature=Base
                      Folder Press FW
                        If False
                          Waypoint WpLmbFwMec: TCP in base x=-30.994 y=682.626 z=386.431 mm, rx=0.3238 ry=3.0539 rz=-0.0115 rad; joints [94.033, -94.235, -107.032, -69.931, 86.424, 196.47] deg; TCP offset x=159 y=-58 z=70 mm, rx=0 ry=0 rz=0 rad
                        Wp := pose_add(WpLmbFwMec,Base_w_correctn)
                        Waypoint Variable (Variable): variable=Wp
                        Timer (action=Reset) variable=T_Timeout
                        Timer (action=Start) variable=T_Timeout
                        Force Frame feature=Joint_6_name; selection=[1, 0, 0, 0, 0, 0]; wrench=[20, 10, -20, 0, 0, 0]; limitsForce=[0.05, 0.01, 0.05, 1.047198, 1.047198, 1.047198]; limitsMotion=[0.1, 0.1, 0.1, 0.349066, 0.349066, 0.349066]
                          Wait Condition expression=Flags[10] or T_Timeout>10 or (DEBUG and T_Timeout>2)
                        Waypoint Variable (Variable): variable=Wp
                  Else 
                    MoveL speed 1000 mm/s, acceleration 3000 mm/s^2 (useActiveTCP=false optimoveEnabled=false optiMoveSpeed=0.3 optiMoveAcceleration=0.09) tcp=t0_Flange; feature=Base
                      Waypoint WpBttnMidp3: motionParameters(blendRadius=0.1); TCP in base x=114.747 y=708.142 z=644.758 mm, rx=0 ry=3.1416 rz=0 rad; joints [94.755, -90.505, -92.903, -86.639, 90.379, 184.947] deg; TCP offset x=0 y=0 z=0 mm, rx=0 ry=0 rz=0 rad
                      Waypoint WpBttnMidp2: motionParameters(blendRadius=0.1); TCP in base x=-296.641 y=583.561 z=625.265 mm, rx=-1.2596 ry=2.878 rz=0 rad; joints [132.275, -84.542, -100.549, -84.955, 90.381, 175.201] deg
                      Waypoint WpBttnMidp1: motionParameters(blendRadius=0.1); TCP in base x=-465.361 y=283.426 z=636.73 mm, rx=-2.2214 ry=2.2214 rz=0 rad; joints [167.185, -73.405, -108.257, -88.385, 90.398, 167.36] deg
                      Waypoint WpHome: TCP in base x=-539.74 y=192.879 z=621.496 mm, rx=3.1416 ry=0 rz=0 rad; joints [177.915, -76.399, -107.627, -86.021, 90.391, 88.106] deg
                    Script: Report(95)
            Folder 2W LMB RW
              If Progress_run()
                If In(ProgExe,[34])
                  Timer (action=Reset) variable=T_Timeout
                  Timer (action=Start) variable=T_Timeout
                  Script: Report(14)
                  Wait Condition expression=Flags[4] or T_Timeout>60 or DEBUG or Abort
                  If Flags[4] or DEBUG
                    MoveL speed 1000 mm/s, acceleration 3000 mm/s^2 (useActiveTCP=false optimoveEnabled=false optiMoveSpeed=0.3 optiMoveAcceleration=0.09) tcp=t4_Finger; feature=Base
                      Folder Press RW
                        If False
                          Waypoint WpLmbRwMec: TCP in base x=-24.827 y=697.185 z=385.645 mm, rx=0.3238 ry=3.0539 rz=-0.0115 rad; joints [93.456, -95.707, -105.506, -69.945, 86.411, 195.892] deg; TCP offset x=159 y=-58 z=70 mm, rx=0 ry=0 rz=0 rad
                        Wp := pose_add(WpLmbRwMec,Base_w_correctn)
                        Waypoint Variable (Variable): variable=Wp
                        Timer (action=Reset) variable=T_Timeout
                        Timer (action=Start) variable=T_Timeout
                        Force Frame feature=Joint_6_name; selection=[1, 0, 0, 0, 0, 0]; wrench=[20, 10, -20, 0, 0, 0]; limitsForce=[0.05, 0.01, 0.05, 1.047198, 1.047198, 1.047198]; limitsMotion=[0.1, 0.1, 0.1, 0.349066, 0.349066, 0.349066]
                          Wait Sleep waitTime=0.5
                        Force Frame feature=Joint_6_name; selection=[1, 0, 0, 0, 0, 0]; wrench=[20, 10, -20, 0, 0, 0]; limitsForce=[0.01, 0.01, 0.05, 1.047198, 1.047198, 1.047198]; limitsMotion=[0.1, 0.1, 0.1, 0.349066, 0.349066, 0.349066]
                          Wait Condition expression=Flags[10] or T_Timeout>10 or (DEBUG and T_Timeout>2)
                        ButtonPos := get_actual_tcp_pose()
                        Waypoint Variable (Variable): variable=Wp
                  Else 
                    MoveL speed 1000 mm/s, acceleration 3000 mm/s^2 (useActiveTCP=false optimoveEnabled=false optiMoveSpeed=0.3 optiMoveAcceleration=0.09) tcp=t0_Flange; feature=Base
                      Waypoint WpBttnMidp3: motionParameters(blendRadius=0.1); TCP in base x=114.747 y=708.142 z=644.758 mm, rx=0 ry=3.1416 rz=0 rad; joints [94.755, -90.505, -92.903, -86.639, 90.379, 184.947] deg; TCP offset x=0 y=0 z=0 mm, rx=0 ry=0 rz=0 rad
                      Waypoint WpBttnMidp2: motionParameters(blendRadius=0.1); TCP in base x=-296.641 y=583.561 z=625.265 mm, rx=-1.2596 ry=2.878 rz=0 rad; joints [132.275, -84.542, -100.549, -84.955, 90.381, 175.201] deg
                      Waypoint WpBttnMidp1: motionParameters(blendRadius=0.1); TCP in base x=-465.361 y=283.426 z=636.73 mm, rx=-2.2214 ry=2.2214 rz=0 rad; joints [167.185, -73.405, -108.257, -88.385, 90.398, 167.36] deg
                      Waypoint WpHome: TCP in base x=-539.74 y=192.879 z=621.496 mm, rx=3.1416 ry=0 rz=0 rad; joints [177.915, -76.399, -107.627, -86.021, 90.391, 88.106] deg
                    Script: Report(95)
            Folder Camera2
              If Progress_run()
                If In(ProgExe,[34])
                  SuppressedNode
                    SetCameraProg := 35
                  MoveL speed 1000 mm/s, acceleration 3000 mm/s^2 (useActiveTCP=false optimoveEnabled=false optiMoveSpeed=0.3 optiMoveAcceleration=0.09) tcp=t0_Flange; feature=Base
                    If False
                      Waypoint WpCamHeightUp: TCP in base x=185.286 y=713.319 z=390.264 mm, rx=0.3312 ry=3.124 rz=0 rad; joints [89.003, -99.18, -110.202, -60.664, 90.284, 191.446] deg
                    Wp := pose_add(WpCamHeightUp,p[0,0,MeasHeight/1000,0,0,0])
                    SuppressedNode
                      Wp := WpCamHeightUp
                    Waypoint Variable (Variable): variable=Wp
                  Call CamAcquire
                  Script: CamData[1]=CamData[1]-MeasHeight/1000
                  Call CamCalculateCorectnPlane
            If Progress_run() and CamCorrectnOK≠ProgExe
              MoveL speed 1000 mm/s, acceleration 3000 mm/s^2 (useActiveTCP=false optimoveEnabled=false optiMoveSpeed=0.3 optiMoveAcceleration=0.09) tcp=t0_Flange; feature=Base
                Waypoint WpBttnMidp3: motionParameters(blendRadius=0.1); TCP in base x=114.747 y=708.142 z=644.758 mm, rx=0 ry=3.1416 rz=0 rad; joints [94.755, -90.505, -92.903, -86.639, 90.379, 184.947] deg; TCP offset x=0 y=0 z=0 mm, rx=0 ry=0 rz=0 rad
                Waypoint WpBttnMidp2: motionParameters(blendRadius=0.1); TCP in base x=-296.641 y=583.561 z=625.265 mm, rx=-1.2596 ry=2.878 rz=0 rad; joints [132.275, -84.542, -100.549, -84.955, 90.381, 175.201] deg
                Waypoint WpBttnMidp1: motionParameters(blendRadius=0.1); TCP in base x=-465.361 y=283.426 z=636.73 mm, rx=-2.2214 ry=2.2214 rz=0 rad; joints [167.185, -73.405, -108.257, -88.385, 90.398, 167.36] deg
                Waypoint WpHome: TCP in base x=-539.74 y=192.879 z=621.496 mm, rx=3.1416 ry=0 rz=0 rad; joints [177.915, -76.399, -107.627, -86.021, 90.391, 88.106] deg
              Script: Report(91)
            Folder Height up
              If Progress_run()
                If In(ProgExe,[34])
                  SetCameraProg := 36
                  Timer (action=Reset) variable=T_Timeout
                  Timer (action=Start) variable=T_Timeout
                  Script: Report(15)
                  Wait Condition expression=Flags[5] or T_Timeout>60 or DEBUG or Abort
                  If Flags[5] or DEBUG
                    MoveL speed 1000 mm/s, acceleration 3000 mm/s^2 (useActiveTCP=false optimoveEnabled=false optiMoveSpeed=0.3 optiMoveAcceleration=0.09) tcp=t4_Finger; feature=Base
                      Folder Press height up
                        If False
                          Waypoint WpHeiUp: TCP in base x=-34.242 y=768.782 z=353.839 mm, rx=-0.3314 ry=-3.1239 rz=-0.0011 rad; joints [92.867, -103.592, -100.979, -65.434, 90.303, 195.294] deg; TCP offset x=159 y=-58 z=70 mm, rx=0 ry=0 rz=0 rad
                        Wp := pose_add(WpHeiUp,Base_w_correctn)
                        SuppressedNode
                          Wp := pose_trans(Wp, p[-0.02,0,0.003,0,0,0])
                        Script: Wp[0]=ButtonPos[0]+0.008
                        Waypoint Variable (Variable): variable=Wp
                        Set NoAction tcp=t4_Finger
                        SuppressedNode
                          Force Frame feature=Joint_6_name; selection=[1, 0, 0, 0, 0, 0]; wrench=[10, 0, 0, 0, 0, 0]; limitsForce=[0.1, 0.15, 0.15, 1.047198, 1.047198, 1.047198]; limitsMotion=[0.1, 0.1, 0.1, 0.349066, 0.349066, 0.349066]
                            Wait Sleep waitTime=0.5
                        SuppressedNode
                          Force Frame feature=Joint_6_name; selection=[1, 0, 0, 0, 0, 0]; wrench=[20, 0, 0, 0, 0, 0]; limitsForce=[0.01, 0.15, 0.15, 1.047198, 1.047198, 1.047198]; limitsMotion=[0.1, 0.1, 0.1, 0.349066, 0.349066, 0.349066]
                            Wait Sleep waitTime=0.5
                        SuppressedNode
                          Wp := pose_trans(P_act, p[-0.002,0,0,0,0,0])
                        SuppressedNode
                          Waypoint Variable (Variable): variable=Wp
                        Timer (action=Reset) variable=T_Timeout
                        Timer (action=Start) variable=T_Timeout
                        Force Frame feature=Base; selection=[0, 1, 1, 0, 0, 0]; wrench=[0, 0, 10, 0, 0, 0]; limitsForce=[0.02, 0.01, 0.05, 1.047198, 1.047198, 1.047198]; limitsMotion=[0.1, 0.1, 0.1, 0.349066, 0.349066, 0.349066]
                          Wait Condition expression=Flags[10] or T_Timeout>10 or (DEBUG and T_Timeout>2)
                        Wp0 := get_actual_tcp_pose()
                        Wp := pose_trans(Wp0, p[-0.02,0,0.02,0,0,0])
                        Waypoint Variable (Variable): variable=Wp
                  Else 
                    MoveL speed 1000 mm/s, acceleration 3000 mm/s^2 (useActiveTCP=false optimoveEnabled=false optiMoveSpeed=0.3 optiMoveAcceleration=0.09) tcp=t0_Flange; feature=Base
                      Waypoint WpBttnMidp3: motionParameters(blendRadius=0.1); TCP in base x=114.747 y=708.142 z=644.758 mm, rx=0 ry=3.1416 rz=0 rad; joints [94.755, -90.505, -92.903, -86.639, 90.379, 184.947] deg; TCP offset x=0 y=0 z=0 mm, rx=0 ry=0 rz=0 rad
                      Waypoint WpBttnMidp2: motionParameters(blendRadius=0.1); TCP in base x=-296.641 y=583.561 z=625.265 mm, rx=-1.2596 ry=2.878 rz=0 rad; joints [132.275, -84.542, -100.549, -84.955, 90.381, 175.201] deg
                      Waypoint WpBttnMidp1: motionParameters(blendRadius=0.1); TCP in base x=-465.361 y=283.426 z=636.73 mm, rx=-2.2214 ry=2.2214 rz=0 rad; joints [167.185, -73.405, -108.257, -88.385, 90.398, 167.36] deg
                      Waypoint WpHome: TCP in base x=-539.74 y=192.879 z=621.496 mm, rx=3.1416 ry=0 rz=0 rad; joints [177.915, -76.399, -107.627, -86.021, 90.391, 88.106] deg
                    Script: Report(95)
            Folder Camera3
              If Progress_run()
                If In(ProgExe,[34])
                  SuppressedNode
                    SetCameraProg := 36
                  MoveL speed 1000 mm/s, acceleration 3000 mm/s^2 (useActiveTCP=false optimoveEnabled=false optiMoveSpeed=0.3 optiMoveAcceleration=0.09) tcp=t0_Flange; feature=Base
                    If False
                      Waypoint WpCamHeightDown: TCP in base x=185.286 y=707.005 z=393.646 mm, rx=-0.3312 ry=-3.1239 rz=0 rad; joints [88.995, -98.468, -110.661, -60.918, 90.286, 191.436] deg
                    Wp := pose_add(WpCamHeightUp,p[0,0,MeasHeight/1000,0,0,0])
                    SuppressedNode
                      Wp := WpCamHeightDown
                    Waypoint Variable (Variable): variable=Wp
                  Call CamAcquire
                  Script: CamData[1]=CamData[1]-MeasHeight/1000
                  Call CamCalculateCorectnPlane
            Folder Height down
              If Progress_run()
                If In(ProgExe,[34])
                  Timer (action=Reset) variable=T_Timeout
                  Timer (action=Start) variable=T_Timeout
                  Script: Report(16)
                  Wait Condition expression=Flags[6] or T_Timeout>60 or DEBUG or Abort
                  If Flags[6] or DEBUG
                    MoveL speed 1000 mm/s, acceleration 3000 mm/s^2 (useActiveTCP=false optimoveEnabled=false optiMoveSpeed=0.3 optiMoveAcceleration=0.09) tcp=t4_Finger; feature=Base
                      Folder Press height down
                        If False
                          Waypoint WpHeiDown: TCP in base x=-33.166 y=771.407 z=382.532 mm, rx=0.1703 ry=3.1369 rz=-0.0001 rad; joints [92.957, -104.254, -97.001, -68.798, 90.311, 189.47] deg; TCP offset x=159 y=-58 z=70 mm, rx=0 ry=0 rz=0 rad
                        Wp := pose_add(WpHeiDown,Base_w_correctn)
                        Script: Wp[0]=ButtonPos[0]+0.008
                        Wp0 := pose_add(Wp,p[0.04,0,0,0,0,0])
                        SuppressedNode
                          Wp := pose_trans(Wp, p[-0.02,0,-0.003,0,0,0])
                        SuppressedNode
                          Wp := pose_trans(WpHeiDown, CamCorrection)
                        SuppressedNode
                          Wp := pose_trans(Wp, p[-0.02,-0.005,0,0,0,0])
                        SuppressedNode
                          Wp := pose_trans(Wp, p[0,0,-0.05,0,0,0])
                        SuppressedNode
                          Waypoint Variable (Variable): variable=Wp
                        SuppressedNode
                          Wp := pose_trans(Wp0, p[0,0,-0.025,0,0,0])
                        Waypoint Variable (Variable): motionParameters(blendRadius=0.03); variable=Wp0
                        Waypoint Variable (Variable): variable=Wp
                        Set NoAction tcp=t4_Finger
                        SuppressedNode
                          Force Frame feature=Joint_6_name; selection=[1, 0, 0, 0, 0, 0]; wrench=[10, 0, 0, 0, 0, 0]; limitsForce=[0.1, 0.15, 0.15, 1.047198, 1.047198, 1.047198]; limitsMotion=[0.1, 0.1, 0.1, 0.349066, 0.349066, 0.349066]
                            Wait Sleep waitTime=0.5
                        SuppressedNode
                          Force Frame feature=Joint_6_name; selection=[1, 0, 0, 0, 0, 0]; wrench=[15, 0, 0, 0, 0, 0]; limitsForce=[0.015, 0.15, 0.15, 1.047198, 1.047198, 1.047198]; limitsMotion=[0.1, 0.1, 0.1, 0.349066, 0.349066, 0.349066]
                            Wait Sleep waitTime=0.5
                        SuppressedNode
                          Wp := pose_trans(P_act, p[-0.004,0,0,0,0,0])
                        SuppressedNode
                          Waypoint Variable (Variable): variable=Wp
                        Timer (action=Reset) variable=T_Timeout
                        Timer (action=Start) variable=T_Timeout
                        Force Frame feature=Base; selection=[0, 1, 1, 0, 0, 0]; wrench=[0, 0, -10, 0, 0, 0]; limitsForce=[0.02, 0.01, 0.05, 1.047198, 1.047198, 1.047198]; limitsMotion=[0.1, 0.1, 0.1, 0.349066, 0.349066, 0.349066]
                          Wait Condition expression=Flags[10] or T_Timeout>10
                        Wp := pose_trans(Wp, p[-0.02,0,-0.02,0,0,0])
                        Waypoint Variable (Variable): variable=Wp
                    Script: Report(7)
                  Else 
                    MoveL speed 1000 mm/s, acceleration 3000 mm/s^2 (useActiveTCP=false optimoveEnabled=false optiMoveSpeed=0.3 optiMoveAcceleration=0.09) tcp=t0_Flange; feature=Base
                      Waypoint WpBttnMidp3: motionParameters(blendRadius=0.1); TCP in base x=114.747 y=708.142 z=644.758 mm, rx=0 ry=3.1416 rz=0 rad; joints [94.755, -90.505, -92.903, -86.639, 90.379, 184.947] deg; TCP offset x=0 y=0 z=0 mm, rx=0 ry=0 rz=0 rad
                      Waypoint WpBttnMidp2: motionParameters(blendRadius=0.1); TCP in base x=-296.641 y=583.561 z=625.265 mm, rx=-1.2596 ry=2.878 rz=0 rad; joints [132.275, -84.542, -100.549, -84.955, 90.381, 175.201] deg
                      Waypoint WpBttnMidp1: motionParameters(blendRadius=0.1); TCP in base x=-465.361 y=283.426 z=636.73 mm, rx=-2.2214 ry=2.2214 rz=0 rad; joints [167.185, -73.405, -108.257, -88.385, 90.398, 167.36] deg
                      Waypoint WpHome: TCP in base x=-539.74 y=192.879 z=621.496 mm, rx=3.1416 ry=0 rz=0 rad; joints [177.915, -76.399, -107.627, -86.021, 90.391, 88.106] deg
                    Script: Report(95)
            If Progress_run()
              MoveL speed 1000 mm/s, acceleration 3000 mm/s^2 (useActiveTCP=false optimoveEnabled=false optiMoveSpeed=0.3 optiMoveAcceleration=0.09) tcp=t0_Flange; feature=Base
                Waypoint WpBttnMidp3: motionParameters(blendRadius=0.1); TCP in base x=114.747 y=708.142 z=644.758 mm, rx=0 ry=3.1416 rz=0 rad; joints [94.755, -90.505, -92.903, -86.639, 90.379, 184.947] deg; TCP offset x=0 y=0 z=0 mm, rx=0 ry=0 rz=0 rad
                Waypoint WpBttnMidp2: motionParameters(blendRadius=0.1); TCP in base x=-296.641 y=583.561 z=625.265 mm, rx=-1.2596 ry=2.878 rz=0 rad; joints [132.275, -84.542, -100.549, -84.955, 90.381, 175.201] deg
                Waypoint WpBttnMidp1: motionParameters(blendRadius=0.1); TCP in base x=-465.361 y=283.426 z=636.73 mm, rx=-2.2214 ry=2.2214 rz=0 rad; joints [167.185, -73.405, -108.257, -88.385, 90.398, 167.36] deg
                Waypoint WpHome: TCP in base x=-539.74 y=192.879 z=621.496 mm, rx=3.1416 ry=0 rz=0 rad; joints [177.915, -76.399, -107.627, -86.021, 90.391, 88.106] deg
              Script: Report(50)
        Folder PushByHandle
          If In(ProgExe,[40])
            Script: Report(1)
            Folder AtHome? [hidden by the author, left out]
            SuppressedNode
              If Progress_run()
                SetCameraProg := 27
                MoveL speed 250 mm/s, acceleration 1200 mm/s^2 (useActiveTCP=false optimoveEnabled=false optiMoveSpeed=0.3 optiMoveAcceleration=0.09) tcp=t0_Flange; feature=Base
                  Waypoint WpBttnMidp1: motionParameters(blendRadius=0.1); TCP in base x=-465.361 y=283.426 z=636.73 mm, rx=-2.2214 ry=2.2214 rz=0 rad; joints [167.185, -73.405, -108.257, -88.385, 90.398, 167.36] deg
                  Waypoint WpBttnMidp2: motionParameters(blendRadius=0.1); TCP in base x=-296.641 y=583.561 z=625.265 mm, rx=-1.2596 ry=2.878 rz=0 rad; joints [132.275, -84.542, -100.549, -84.955, 90.381, 175.201] deg
                  Waypoint WpBttnMidp3: motionParameters(blendRadius=0.1); TCP in base x=114.747 y=708.142 z=644.758 mm, rx=0 ry=3.1416 rz=0 rad; joints [94.755, -90.505, -92.903, -86.639, 90.379, 184.947] deg; TCP offset x=0 y=0 z=0 mm, rx=0 ry=0 rz=0 rad
                  Waypoint WpCamLMB: TCP in base x=186.376 y=644.645 z=421.712 mm, rx=0.3238 ry=3.0539 rz=-0.0115 rad; joints [89.517, -91.476, -115.043, -64.369, 86.327, 191.973] deg
                Call CamAcquire
                CamCorrection := p[0,CamData[0],CamData[1],0,0,0]
            SuppressedNode
              If Progress_run() and CamCorrectnOK≠ProgExe
                MoveL speed 250 mm/s, acceleration 1200 mm/s^2 (useActiveTCP=false optimoveEnabled=false optiMoveSpeed=0.3 optiMoveAcceleration=0.09) tcp=t0_Flange; feature=Base
                  Waypoint WpBttnMidp3: motionParameters(blendRadius=0.1); TCP in base x=114.747 y=708.142 z=644.758 mm, rx=0 ry=3.1416 rz=0 rad; joints [94.755, -90.505, -92.903, -86.639, 90.379, 184.947] deg; TCP offset x=0 y=0 z=0 mm, rx=0 ry=0 rz=0 rad
                  Waypoint WpBttnMidp2: motionParameters(blendRadius=0.1); TCP in base x=-296.641 y=583.561 z=625.265 mm, rx=-1.2596 ry=2.878 rz=0 rad; joints [132.275, -84.542, -100.549, -84.955, 90.381, 175.201] deg
                  Waypoint WpBttnMidp1: motionParameters(blendRadius=0.1); TCP in base x=-465.361 y=283.426 z=636.73 mm, rx=-2.2214 ry=2.2214 rz=0 rad; joints [167.185, -73.405, -108.257, -88.385, 90.398, 167.36] deg
                  Waypoint WpHome: TCP in base x=-539.74 y=192.879 z=621.496 mm, rx=3.1416 ry=0 rz=0 rad; joints [177.915, -76.399, -107.627, -86.021, 90.391, 88.106] deg
                Script: Report(91)
            If Progress_run() and  not AdapterDocked
              Script: Report(94)
            If Progress_run()
              PusherReturn := False
              Set DigitalOutput pin=Do_PusherReturn; digitalValue=0
              Set DigitalOutput pin=Do_PusherWork; digitalValue=1
              Wait Condition expression=PusherPosStable and PusherPosDev>-20
              Set DigitalOutput pin=Do_PusherWork; digitalValue=0
              Call GripperOpen
              Set NoAction tcp=t2_Gripper
              MoveL speed 1000 mm/s, acceleration 3000 mm/s^2 (useActiveTCP=false optimoveEnabled=false optiMoveSpeed=0.3 optiMoveAcceleration=0.09) tcp=t2_Gripper; feature=Base
                Waypoint WpHandle0: motionParameters(blendRadius=0.05); TCP in base x=-455.859 y=509.138 z=225.989 mm, rx=3.1416 ry=0 rz=0 rad; joints [170.787, -84.178, -136.861, -49.009, 90.24, 81.174] deg; TCP offset x=0 y=-260 z=74 mm, rx=0 ry=0 rz=0 rad
                Waypoint WpHandle: TCP in base x=-329.851 y=672.326 z=234.484 mm, rx=3.1416 ry=0 rz=0 rad; joints [147.777, -84.364, -135.583, -50.1, 90.246, 58.16] deg
                Force Frame feature=Joint_6_name; selection=[0, 1, 0, 0, 0, 0]; wrench=[0, -10, 0, 0, 0, 0]; limitsForce=[0.15, 0.05, 0.15, 1.047198, 1.047198, 1.047198]; limitsMotion=[0.1, 0.1, 0.1, 0.349066, 0.349066, 0.349066]
                  Wait Sleep waitTime=1
                Force Frame feature=Joint_6_name; selection=[0, 1, 1, 0, 0, 0]; wrench=[0, -10, -80, 0, 0, 0]; limitsForce=[0.15, 0.05, 0.05, 1.047198, 1.047198, 1.047198]; limitsMotion=[0.1, 0.1, 0.1, 0.349066, 0.349066, 0.349066]
                  Wait Sleep waitTime=1
                Force Frame feature=Joint_6_name; selection=[0, 1, 1, 0, 0, 0]; wrench=[0, -30, -80, 0, 0, 0]; limitsForce=[0.15, 0.5, 0.05, 1.047198, 1.047198, 1.047198]; limitsMotion=[0.1, 0.1, 0.1, 0.349066, 0.349066, 0.349066]
                  Wait Sleep waitTime=0.2
                  Set DigitalOutput pin=Do_PusherReturn; digitalValue=0
                  Set DigitalOutput pin=Do_PusherWork; digitalValue=1
                  Wait AnalogInput pin=analog_in[0]; analogComparison=0; analogValue=8.9
                  Wait Sleep waitTime=2
                  Set DigitalOutput pin=Do_PusherWork; digitalValue=0
                PusherReturn := True
                Waypoint WpOffHandle (Relative): relativeFromPosition TCP in base x=-352.096 y=769.969 z=292.34 mm, rx=3.1371 ry=-0.0001 rz=0.0084 rad; joints [140.822, -89.589, -123.274, -57.586, 90.286, 51.179] deg; TCP in base x=-351.703 y=761.028 z=222.838 mm, rx=3.1371 ry=-0.0002 rz=0.0084 rad; joints [141.47, -93.676, -127.767, -49.003, 90.241, 51.867] deg
                Waypoint WpHandle0: TCP in base x=-455.859 y=509.138 z=225.989 mm, rx=3.1416 ry=0 rz=0 rad; joints [170.787, -84.178, -136.861, -49.009, 90.24, 81.174] deg
              MoveL speed 1000 mm/s, acceleration 3000 mm/s^2 (useActiveTCP=false optimoveEnabled=false optiMoveSpeed=0.3 optiMoveAcceleration=0.09) tcp=t0_Flange; feature=Base
                Waypoint WpHome: TCP in base x=-539.74 y=192.879 z=621.496 mm, rx=3.1416 ry=0 rz=0 rad; joints [177.915, -76.399, -107.627, -86.021, 90.391, 88.106] deg
              Script: Report(50)
        Folder Tilt manual adjust
          If In(ProgExe,[42])
            Script: Report(1)
            Folder AtHome? [hidden by the author, left out]
            If Progress_run() and  not AdapterDocked
              Script: Report(94)
            If Progress_run()
              Set NoAction tcp=t2_Gripper
              ''
              If InRange(Tilt_PV-CMD_Tilt_SP,-60,60)
                'Laser value in range'
                MaxTiltPumps := 10
                If InRange(Tilt_PV-CMD_Tilt_SP,-60,-3)
                  'Tilt too high'
                  Call GripperClose
                  MoveJ speed 120 deg/s, acceleration 500 deg/s^2 (useActiveTCP=false positionType=JointAngles optimoveEnabled=false optiMoveSpeed=0.3 optiMoveAcceleration=0.09) tcp=t2_Gripper; feature=Base
                    Waypoint WpTilt0: motionParameters(blendRadius=0.05); TCP in base x=-583.368 y=339.327 z=316.361 mm, rx=1.6182 ry=-0.1906 rz=-1.3026 rad; joints [156.708, -75.754, -120.579, -153.057, 211.083, -30.966] deg; TCP offset x=0 y=-260 z=74 mm, rx=0 ry=0 rz=0 rad
                    Waypoint WpTilt1: motionParameters(blendRadius=0.05); TCP in base x=-466.465 y=329.412 z=219.468 mm, rx=1.2093 ry=-1.2091 rz=-1.2092 rad; joints [153.941, -75.671, -122.269, -161.849, 244.19, 0.382] deg
                    Waypoint WpTiltDown: TCP in base x=-481.518 y=636.8 z=214.526 mm, rx=1.5185 ry=-0.974 rz=-1.5185 rad; joints [135.681, -94.646, -108.169, -156.834, 225.958, -24.187] deg
                    Force Frame feature=Joint_6_name; selection=[1, 1, 0, 0, 0, 0]; wrench=[-15, 0, 0, 0, 0, 0]; limitsForce=[0.1, 0.15, 0.15, 1.047198, 1.047198, 1.047198]; limitsMotion=[0.1, 0.1, 0.1, 0.349066, 0.349066, 0.349066]
                      Wait Sleep waitTime=1
                    Wp := P_act
                    Loop While (checkContinuously=false) expression=InRange(Tilt_PV-CMD_Tilt_SP,-60,-5) and MaxTiltPumps>0
                      Force Frame feature=Joint_6_name; selection=[1, 1, 0, 0, 0, 0]; wrench=[-10, -100, 0, 0, 0, 0]; limitsForce=[0.15, 0.1, 0.15, 1.047198, 1.047198, 1.047198]; limitsMotion=[0.1, 0.1, 0.1, 0.349066, 0.349066, 0.349066]
                        Wait Sleep waitTime=1.5
                      Waypoint Variable (Variable): variable=Wp
                      MaxTiltPumps := MaxTiltPumps-1
                    Waypoint WpTiltDown: motionParameters(blendRadius=0.05); TCP in base x=-481.518 y=636.8 z=214.526 mm, rx=1.5185 ry=-0.974 rz=-1.5185 rad; joints [135.681, -94.646, -108.169, -156.834, 225.958, -24.187] deg
                    Waypoint WpTilt1: motionParameters(blendRadius=0.05); TCP in base x=-466.465 y=329.412 z=219.468 mm, rx=1.2093 ry=-1.2091 rz=-1.2092 rad; joints [153.941, -75.671, -122.269, -161.849, 244.19, 0.382] deg
                    Waypoint WpTilt0: TCP in base x=-583.368 y=339.327 z=316.361 mm, rx=1.6182 ry=-0.1906 rz=-1.3026 rad; joints [156.708, -75.754, -120.579, -153.057, 211.083, -30.966] deg
                  MoveJ speed 120 deg/s, acceleration 500 deg/s^2 (useActiveTCP=false positionType=JointAngles optimoveEnabled=false optiMoveSpeed=0.3 optiMoveAcceleration=0.09) tcp=t0_Flange; feature=Base
                    Waypoint WpHome: TCP in base x=-539.74 y=192.879 z=621.496 mm, rx=3.1416 ry=0 rz=0 rad; joints [177.915, -76.399, -107.627, -86.021, 90.391, 88.106] deg
                ElseIf InRange(Tilt_PV-CMD_Tilt_SP,3,60)
                  'Tilt too low'
                  Call GripperClose
                  MoveJ speed 120 deg/s, acceleration 500 deg/s^2 (useActiveTCP=false positionType=JointAngles optimoveEnabled=false optiMoveSpeed=0.3 optiMoveAcceleration=0.09) tcp=t2_Gripper; feature=Base
                    Waypoint WpTilt0: motionParameters(blendRadius=0.05); TCP in base x=-583.368 y=339.327 z=316.361 mm, rx=1.6182 ry=-0.1906 rz=-1.3026 rad; joints [156.708, -75.754, -120.579, -153.057, 211.083, -30.966] deg; TCP offset x=0 y=-260 z=74 mm, rx=0 ry=0 rz=0 rad
                    Waypoint WpTilt1: motionParameters(blendRadius=0.05); TCP in base x=-466.465 y=329.412 z=219.468 mm, rx=1.2093 ry=-1.2091 rz=-1.2092 rad; joints [153.941, -75.671, -122.269, -161.849, 244.19, 0.382] deg
                    Waypoint WpTiltUp: TCP in base x=-484.61 y=613.687 z=229.929 mm, rx=1.3457 ry=-1.1148 rz=-1.3455 rad; joints [133.402, -96.666, -102.216, -160.73, 223.658, -10.225] deg
                    Force Frame feature=Joint_6_name; selection=[1, 1, 0, 0, 0, 0]; wrench=[-15, 0, 0, 0, 0, 0]; limitsForce=[0.1, 0.15, 0.15, 1.047198, 1.047198, 1.047198]; limitsMotion=[0.1, 0.1, 0.1, 0.349066, 0.349066, 0.349066]
                      Wait Sleep waitTime=1
                    Wp := P_act
                    Loop While (checkContinuously=false) expression=InRange(Tilt_PV-CMD_Tilt_SP,5,60) and MaxTiltPumps>0
                      Force Frame feature=Joint_6_name; selection=[1, 1, 0, 0, 0, 0]; wrench=[-10, 100, 0, 0, 0, 0]; limitsForce=[0.15, 0.1, 0.15, 1.047198, 1.047198, 1.047198]; limitsMotion=[0.1, 0.1, 0.1, 0.349066, 0.349066, 0.349066]
                        Wait Sleep waitTime=1.5
                      Waypoint Variable (Variable): variable=Wp
                      MaxTiltPumps := MaxTiltPumps-1
                    Waypoint WpTiltUp: motionParameters(blendRadius=0.05); TCP in base x=-484.61 y=613.687 z=229.929 mm, rx=1.3457 ry=-1.1148 rz=-1.3455 rad; joints [133.402, -96.666, -102.216, -160.73, 223.658, -10.225] deg
                    Waypoint WpTilt1: motionParameters(blendRadius=0.05); TCP in base x=-466.465 y=329.412 z=219.468 mm, rx=1.2093 ry=-1.2091 rz=-1.2092 rad; joints [153.941, -75.671, -122.269, -161.849, 244.19, 0.382] deg
                    Waypoint WpTilt0: motionParameters(blendRadius=0.05); TCP in base x=-583.368 y=339.327 z=316.361 mm, rx=1.6182 ry=-0.1906 rz=-1.3026 rad; joints [156.708, -75.754, -120.579, -153.057, 211.083, -30.966] deg
                    Waypoint WpHome: TCP in base x=-539.74 y=192.879 z=621.496 mm, rx=3.1416 ry=0 rz=0 rad; joints [177.915, -76.399, -107.627, -86.021, 90.391, 88.106] deg
              Else 
                Script: Report(93)
              Script: Report(50)
        Folder Program finished
          ProgDn := ProgExe
          ProgExe := 0
      Folder Parking
        If Parking≟10 or ProgExe≟1011
          Wait Condition expression=EvtDock≤0
          If AtHomePos
            MoveJ speed 120 deg/s, acceleration 500 deg/s^2 (useActiveTCP=true positionType=JointAngles optimoveEnabled=false optiMoveSpeed=0.3 optiMoveAcceleration=0.09) feature=Base
              Waypoint WpPark: TCP in base x=153.666 y=469.873 z=822.74 mm, rx=-0.0357 ry=3.1413 rz=-0.0002 rad; joints [92.418, -70.926, -90.975, -108.153, 90.407, 181.161] deg
              STS_Reservation := 0
          Parking := 0
          If DEBUG
            ProgExe := 0
        If Parking≟1 or ProgExe≟1001
          If AtParkPos
            MoveJ speed 120 deg/s, acceleration 500 deg/s^2 (useActiveTCP=true positionType=JointAngles optimoveEnabled=false optiMoveSpeed=0.3 optiMoveAcceleration=0.09) feature=Base
              Waypoint WpHome: TCP in base x=-539.74 y=192.879 z=621.496 mm, rx=3.1416 ry=0 rz=0 rad; joints [177.915, -76.399, -107.627, -86.021, 90.391, 88.106] deg
              STS_Reservation := 1
            Parking := 0
            If DEBUG
              ProgExe := 0
  Script: sync()
Thread Thread_1 (runOnlyOnce=false)
  Folder Continuous calculations
    Folder get live force and tcp pos
      P_act := get_actual_tcp_pose()
      V_act := get_actual_tcp_speed()
      V_act_norm := norm(V_act)
      ToolForce := norm(get_tcp_force())
      P_Flange := get_actual_tool_flange_pose()
      D_rel := pose_sub(P_act, P_ini)
      AtHomePos := pose_dist(P_Flange, WpHome)<0.005
      AtParkPos := pose_dist(P_Flange, WpPark)<0.005
      AdapterDocked := Di_Docked
      Tilt_PV := (Ai_LaserTilt*100+505)*0.1+Tilt_PV*0.9
      Folder Calculate actual offset in tool frame
        If ProgExe≟15
          TempWp := pose_sub(WpBuckleSpa1,Base_w_correctn)
          BklToolDist := pose_trans(pose_inv(TempWp), P_act)
        If ProgExe≟16
          TempWp := pose_sub(WpBuckleSpa3,Base_w_correctn)
          BklToolDist := pose_trans(pose_inv(TempWp), P_act)
      Folder InterlockOutput
        If P_Flange[1]>-0.45
          Set DigitalOutput pin=Do_SafePosition; digitalValue=1
        ElseIf P_Flange[0]>0
          Set DigitalOutput pin=Do_SafePosition; digitalValue=1
        Else 
          Set DigitalOutput pin=Do_SafePosition; digitalValue=0
    Folder Modbus mapping
      Folder Heartbeat
        Timer (action=Start) variable(name=T_Heartbeat)
        If T_Heartbeat≥1
          Timer (action=Reset) variable=T_Heartbeat
          If STS_Heartbeat
            STS_Heartbeat := False
          Else 
            STS_Heartbeat := True
      Folder Safe position
        STS_Safe := True
        If pose_dist(P_act,WpBuckleSpa1)<0.2
          STS_Safe := False
        If pose_dist(P_act,WpConnSpa1EL)<0.08
          STS_Safe := False
        If pose_dist(P_act,WpHandle)<0.08
          STS_Safe := False
        If pose_dist(P_act,WpHeiUp)<0.08
          STS_Safe := False
        If pose_dist(P_act,WpLmbFwEL)<0.08
          STS_Safe := False
        If pose_dist(P_act,WpUnplug1_3)<0.08
          STS_Safe := False
        If pose_dist(P_act,WpUnplg1_3M)<0.08
          STS_Safe := False
      Folder Outputs
        Script: write_port_register(129,STS_Progress)
        Script: write_port_register(131,STS_Reservation)
        Script: write_port_register(134,binary_list_to_integer([digital_in[0], False ,config_in[0],STS_Heartbeat,STS_Safe, False ]))
      Folder Inputs
        CMD_Reserve_i1 := read_port_register(160)
        CMD_Timeout_i1 := read_port_register(162)
        CMD_Program_i1 := read_port_register(164)
        CMD_Tilt_SP := read_port_register(166)
        CMD_Flags_i1 := read_port_register(170)
        CMD_Heartbt_i1 := read_port_register(180)
      Folder Generate flags
        Flags := integer_to_binary_list(CMD_Flags_i1)
    Folder Speed
      Timer (action=Start) variable(name=T_SpeedSet)
      If T_SpeedSet>2 and  not DEBUG
        Script: socket_send_string("set speed")
        Script: socket_send_string(1.0)
        Script: socket_send_byte(10)
        Timer (action=Reset) variable=T_SpeedSet
    Wait Sleep waitTime=0.01
  Folder ReservationControl
    If STS_Reservation≟0 and ProgExe≟0
      If CMD_Reserve_i1≟1
        'request reservation'
        If AtHomePos or AdapterReady
          STS_Reservation := 1
        Else 
          Parking := 1
    'Timeout reservation - station keeps reservation for a while to prevent other app stealing the process'
    'Timeout is configurable, so application can control how long to keep robot before letting other app'
    If STS_Progress≟0 and STS_Reservation≠0
      If STS_Reservation≟1 and CMD_Reserve_i1≟1
        'nop'
      Else 
        T_KeepReservtn := CMD_Timeout_i1
        Timer (action=Start) variable(name=tim_Unreserve)
        If tim_Unreserve>T_KeepReservtn
          STS_Reservation := 0
          Timer (action=Stop) variable=tim_Unreserve
    Else 
      Timer (action=Stop) variable=tim_Unreserve
      Timer (action=Reset) variable=tim_Unreserve
    'Force release reservation from app - in case of intervetion'
    If STS_Progress≟0 and In(STS_Reservation,[0,1]) and In(CMD_Reserve_i1,[98,99]) and  not DEBUG
      If AtHomePos
        Parking := 10
      If AtParkPos
        STS_Reservation := 0
      If CMD_Reserve_i1≟99 and  not Mute
        Set DigitalOutput pin=Do_Blue; digitalValue=1
        Set DigitalOutput pin=Do_Horn; digitalValue=1
    Wait Sleep waitTime=0.01
  Folder Program control
    'Start new Prog / Confirm Prog Running'
    If STS_Progress≟0 and ProgExe≟0  and  not Abort and  not DEBUG
      If InRange(CMD_Program_i1,10,49) and STS_Reservation≟1
        ProgExe := CMD_Program_i1
        T_KeepReservtn := CMD_Timeout_i1
        Script: Report(0)
    'Ack results - get ready for new prg'
    If ProgExe≟0 and Progress_finished()
      If CMD_Program_i1≠ProgDn
        STS_Progress := 0
  Folder Pusher Control
    If PusherReturn and NormalMode
      Set DigitalOutput pin=Do_PusherReturn; digitalValue=1
      Set DigitalOutput pin=Do_PusherWork; digitalValue=0
      Timer (action=Start) variable(name=T_Pusher)
      If T_Pusher>20 or Di_Pusher_Bp
        Set DigitalOutput pin=Do_PusherReturn; digitalValue=0
        PusherReturn := False
    Else 
      Timer (action=Stop) variable=T_Pusher
      Timer (action=Reset) variable=T_Pusher
    If not NormalMode
      Set DigitalOutput pin=Do_PusherReturn; digitalValue=0
      Set DigitalOutput pin=Do_PusherWork; digitalValue=0
    If Flags[11] and NormalMode
      'Activate pusher in advance'
      Set DigitalOutput pin=Do_PusherReturn; digitalValue=0
      Set DigitalOutput pin=Do_PusherWork; digitalValue=1
    PusherPos := Calibrate(Ai_Pusher,1,8,260,385)
    PusherPosFt := PusherPos*0.2+PusherPosFt*0.8
    PusherPosStable := InRange(PusherPosFt-PusherPos,-1,1) and PusherPosFt>265
  Folder Operator call deactivation
    If Do_Blue or Do_Horn
      Timer (action=Start) variable(name=T_Call)
      If not  NormalMode and T_Call>4
        Set DigitalOutput pin=Do_Blue; digitalValue=0
        Set DigitalOutput pin=Do_Horn; digitalValue=0
        Mute := True
    Else 
      Timer (action=Stop) variable=T_Call
      Timer (action=Reset) variable=T_Call
  Folder Abort
    If Flags[14]
      Abort := True
    If AtHomePos or AtParkPos
      Abort := False
    If Abort
      If AdapterReady
        EvtDock := 1
  Wait Sleep waitTime=0.01
SubProgram WaitForNormalMode [hidden by the author, left out]
SubProgram  [hidden by the author, left out]
SubProgram  [hidden by the author, left out]
SubProgram  [hidden by the author, left out]
SubProgram  [hidden by the author, left out]
Event  expression=SetCameraProg>0
  Folder Set program to camera in advance
    Set DigitalOutput pin=CnxDO_Trig; digitalValue=0
    Set DigitalOutput pin=CnxDO_TrigEn; digitalValue=1
    Script: modbus_delete_signal("CnxAO_Program")
    Script: modbus_add_signal("192.168.1.101", 255, 2001, 16, "CnxAO_Program", True ,1)
    Script: modbus_set_output_register("CnxAO_Program",SetCameraProg, False )
    Wait Sleep waitTime=0.2
    Set DigitalOutput pin=CnxDO_SetUsrDta; digitalValue=1
    Wait DigitalInput pin=CnxDi_UsrDtaAck; digitalValue=1
    Set DigitalOutput pin=CnxDO_SetUsrDta; digitalValue=0
    Set DigitalOutput pin=CnxDO_SoftEvt0; digitalValue=1
    Wait DigitalInput pin=CnxDI_Evt0Ack; digitalValue=1
    Set DigitalOutput pin=CnxDO_SoftEvt0; digitalValue=0
    Timer (action=Reset) variable=CamTimeout
    Timer (action=Start) variable=CamTimeout
    Wait Condition expression=CnxAI_Program≟SetCameraProg or CamTimeout>3
    If CnxAI_Program≠SetCameraProg
      Folder For the first time it needs trigger when going online
        Set DigitalOutput pin=CnxDO_Trig; digitalValue=1
        Wait Sleep waitTime=1
        Set DigitalOutput pin=CnxDO_Trig; digitalValue=0
        Script: textmsg("extra cam trigger on program set")
      If CnxAI_Program≠SetCameraProg
        SuppressedNode
          Popup Error (haltProgram=false message=Error: camera program not set inputType=Text)
      Else 
        Wait Sleep waitTime=0.5
        SetCameraProg := 0
    Else 
      Wait Sleep waitTime=0.5
      SetCameraProg := 0
  If SetCameraProg>0
    'repeat on fail'
    Wait Sleep waitTime=3
    Folder Set program to camera in advance
      Set DigitalOutput pin=CnxDO_Trig; digitalValue=0
      Set DigitalOutput pin=CnxDO_TrigEn; digitalValue=1
      Script: modbus_delete_signal("CnxAO_Program")
      Script: modbus_add_signal("192.168.1.101", 255, 2001, 16, "CnxAO_Program", True ,1)
      Script: modbus_set_output_register("CnxAO_Program",SetCameraProg, False )
      Wait Sleep waitTime=0.2
      Set DigitalOutput pin=CnxDO_SetUsrDta; digitalValue=1
      Wait DigitalInput pin=CnxDi_UsrDtaAck; digitalValue=1
      Set DigitalOutput pin=CnxDO_SetUsrDta; digitalValue=0
      Set DigitalOutput pin=CnxDO_SoftEvt0; digitalValue=1
      Wait DigitalInput pin=CnxDI_Evt0Ack; digitalValue=1
      Set DigitalOutput pin=CnxDO_SoftEvt0; digitalValue=0
      Timer (action=Reset) variable=CamTimeout
      Timer (action=Start) variable=CamTimeout
      Wait Condition expression=CnxAI_Program≟SetCameraProg or CamTimeout>3
      If CnxAI_Program≠SetCameraProg
        Folder For the first time it needs trigger when going online
          Set DigitalOutput pin=CnxDO_Trig; digitalValue=1
          Wait Sleep waitTime=1
          Set DigitalOutput pin=CnxDO_Trig; digitalValue=0
          Script: textmsg("extra cam trigger on program set")
        If CnxAI_Program≠SetCameraProg
          SuppressedNode
            Popup Error (haltProgram=false message=Error: camera program not set inputType=Text)
        Else 
          Wait Sleep waitTime=0.5
          SetCameraProg := 0
      Else 
        Wait Sleep waitTime=0.5
        SetCameraProg := 0
  If SetCameraProg>0
    'repeat on fail'
    Wait Sleep waitTime=3
    Folder Set program to camera in advance
      Set DigitalOutput pin=CnxDO_Trig; digitalValue=0
      Set DigitalOutput pin=CnxDO_TrigEn; digitalValue=1
      Script: modbus_delete_signal("CnxAO_Program")
      Script: modbus_add_signal("192.168.1.101", 255, 2001, 16, "CnxAO_Program", True ,1)
      Script: modbus_set_output_register("CnxAO_Program",SetCameraProg, False )
      Wait Sleep waitTime=0.2
      Set DigitalOutput pin=CnxDO_SetUsrDta; digitalValue=1
      Wait DigitalInput pin=CnxDi_UsrDtaAck; digitalValue=1
      Set DigitalOutput pin=CnxDO_SetUsrDta; digitalValue=0
      Set DigitalOutput pin=CnxDO_SoftEvt0; digitalValue=1
      Wait DigitalInput pin=CnxDI_Evt0Ack; digitalValue=1
      Set DigitalOutput pin=CnxDO_SoftEvt0; digitalValue=0
      Timer (action=Reset) variable=CamTimeout
      Timer (action=Start) variable=CamTimeout
      Wait Condition expression=CnxAI_Program≟SetCameraProg or CamTimeout>3
      If CnxAI_Program≠SetCameraProg
        Folder For the first time it needs trigger when going online
          Set DigitalOutput pin=CnxDO_Trig; digitalValue=1
          Wait Sleep waitTime=1
          Set DigitalOutput pin=CnxDO_Trig; digitalValue=0
          Script: textmsg("extra cam trigger on program set")
        If CnxAI_Program≠SetCameraProg
          SuppressedNode
            Popup Error (haltProgram=false message=Error: camera program not set inputType=Text)
        Else 
          Wait Sleep waitTime=0.5
          SetCameraProg := 0
      Else 
        Wait Sleep waitTime=0.5
        SetCameraProg := 0
  If SetCameraProg>0
    Popup Error (haltProgram=false message=Error: camera program not set inputType=Text)
SubProgram -> CamAcquire
SubProgram -> CamCalculateCorectnPlane
Event  expression=EvtDock>0
  Folder Dock
    MoveL speed 1000 mm/s, acceleration 3000 mm/s^2 (useActiveTCP=false optimoveEnabled=false optiMoveSpeed=0.3 optiMoveAcceleration=0.09) tcp=t2_Gripper; feature=Base
      If EvtDock≟2
        Folder Force mvts
          Set NoAction tcp=t2_Gripper
          Wp0 := P_act
          Force Frame feature=Joint_6_name; selection=[0, 1, 0, 0, 0, 0]; wrench=[0, -20, 0, 0, 0, 0]; limitsForce=[0.15, 0.1, 0.15, 1.047198, 1.047198, 1.047198]; limitsMotion=[0.1, 0.1, 0.1, 0.349066, 0.349066, 0.349066]
            Wait Sleep waitTime=1
          Force Frame feature=Joint_6_name; selection=[1, 0, 1, 0, 0, 0]; wrench=[0, -10, 0, 0, 0, 0]; limitsForce=[0.15, 0.05, 0.1, 1.047198, 1.047198, 1.047198]; limitsMotion=[0.1, 0.1, 0.1, 0.349066, 0.349066, 0.349066]
            Wait Sleep waitTime=0.2
            Call GripperClose
            Wait Sleep waitTime=0.2
          If timer_Gripper>3
            Call GripperOpen
            MoveL speed 500 mm/s, acceleration 1200 mm/s^2 (useActiveTCP=true optimoveEnabled=false optiMoveSpeed=0.3 optiMoveAcceleration=0.09) feature=Base
              Waypoint Variable (Variable): variable=Wp0
            Force Frame feature=Joint_6_name; selection=[0, 1, 0, 0, 0, 0]; wrench=[0, -20, 0, 0, 0, 0]; limitsForce=[0.15, 0.1, 0.15, 1.047198, 1.047198, 1.047198]; limitsMotion=[0.1, 0.1, 0.1, 0.349066, 0.349066, 0.349066]
              Wait Sleep waitTime=1
            Force Frame feature=Joint_6_name; selection=[1, 0, 1, 0, 0, 0]; wrench=[0, -10, 0, 0, 0, 0]; limitsForce=[0.15, 0.05, 0.1, 1.047198, 1.047198, 1.047198]; limitsMotion=[0.1, 0.1, 0.1, 0.349066, 0.349066, 0.349066]
              Wait Sleep waitTime=0.2
              Call GripperClose
              Wait Sleep waitTime=0.2
          If timer_Gripper>3
            Call GripperOpen
            MoveL speed 500 mm/s, acceleration 1200 mm/s^2 (useActiveTCP=true optimoveEnabled=false optiMoveSpeed=0.3 optiMoveAcceleration=0.09) feature=Base
              Waypoint Variable (Variable): variable=Wp0
              EvtDock := -97
          If EvtDock≟2
            MoveDirectionNode (selectedDirection=YPlus) feature=Joint_6_name
              Until DISTANCE (allowActions=false deceleration=3 distanceNodeType=BLEND) Distance=0.05; motionParameters(blendRadius=0.04)
      If EvtDock>0
        Wp := pose_trans(WpDock, p[0,0.25,0.1,0,0,0])
        Script: Report(40)
        Waypoint Variable (Variable): motionParameters(blendRadius=0.05); variable=Wp
        Wp := pose_trans(WpDock, p[0,0.25,0,0,0,0])
        Waypoint Variable (Variable): motionParameters(blendRadius=0.05); variable=Wp
        Waypoint WpDock referenceName=WpDock: TCP in base x=-876.296 y=277.871 z=78.699 mm, rx=1.8725 ry=1.8725 rz=0.5904 rad; joints [172.393, -110.839, -101.123, -92.857, 86.047, -6.096] deg; TCP offset x=0 y=-260 z=74 mm, rx=0 ry=0 rz=0 rad
        Call GripperOpen
        Waypoint Variable (Variable): variable=Wp
        MoveL speed 1000 mm/s, acceleration 3000 mm/s^2 (useActiveTCP=false optimoveEnabled=false optiMoveSpeed=0.3 optiMoveAcceleration=0.09) tcp=t0_Flange; feature=Base
          Waypoint WpHome: TCP in base x=-539.74 y=192.879 z=621.496 mm, rx=3.1416 ry=0 rz=0 rad; joints [177.915, -76.399, -107.627, -86.021, 90.391, 88.106] deg
        EvtDock := 0
    AdapterReady := False
Event  expression=EvtBeep
  Loop While (checkContinuously=false) expression=EvtBeep
    Set DigitalOutput pin=Do_Horn; digitalValue=1
    Set DigitalOutput pin=Do_Blue; digitalValue=1
    Wait Sleep waitTime=0.5
    Set DigitalOutput pin=Do_Horn; digitalValue=0
    Set DigitalOutput pin=Do_Blue; digitalValue=0
    Wait Sleep waitTime=5
SubProgram GripperOpen [hidden by the author, left out]
SubProgram GripperOpenQuick [hidden by the author, left out]
SubProgram GripperClose [hidden by the author, left out]
SubProgram CamAcquire (keepSynchronizedWithDisk=false)
  Folder Trig camera and process data
    Folder Init
      CamCorrectnOK := 0
      CamRetry := 0
    Wait Condition expression=SetCameraProg≟0
    Loop While (checkContinuously=false) expression=CamRetry<3
      Folder Trig
        CnxCounter := CnxAI_Counter
        Set DigitalOutput pin=CnxDO_Trig; digitalValue=1
        Timer (action=Reset) variable(name=CamTimeout)
        Timer (action=Start) variable=CamTimeout
        Wait Condition expression=CamTimeout>1 or CnxAI_Counter≠CnxCounter
        Set DigitalOutput pin=CnxDO_Trig; digitalValue=0
        Wait Sleep waitTime=0.2
        If CnxAI_Result≥100 and CnxAI_Counter≠CnxCounter
          CamRetry := 100
        Else 
          Wait Sleep waitTime=1
          CamRetry := CamRetry+1
    Folder New data validation
      If CamRetry≟100
        CamCorrectnOK := ProgExe
      Else 
        CamCorrectnOK := 0
      CamData := [(CnxAI_ResultX-30000)/10000,(CnxAI_ResultY-30000)/10000,d2r((CnxAI_ResultR-30000)/10)]
      SuppressedNode
        If CamData[1]>0.03
          Err_state := 103
      SuppressedNode
        If CamData[1]<-0.03
          Err_state := 104
      SuppressedNode
        If CamData[2]>15
          Err_state := 105
      SuppressedNode
        If CamData[2]<-15
          Err_state := 106
SubProgram GripperCloseQuick [hidden by the author, left out]
SubProgram CamCalculateCorectnPlane (keepSynchronizedWithDisk=false)
  Folder Folder
    Set NoAction tcp=t0_Flange
    Script: sync()
    P_act := get_actual_tcp_pose()
    CamCorrection := p[0,CamData[0],CamData[1],0,0,0]
    CamOffset := pose_trans(P_act,CamCorrection)
    Base_w_correctn := pose_sub(CamOffset, P_act)
